(* IEC 61131-3 sources: codesys_asrs/Project_ASRS_CodeSYS, 27 files *)

(* ---- 00_DUT_UDT_MOULE.st ---- *)
// ================================================================
// 00_DUT_UDT_MOULE.st  —  Type utilisateur AS/RS QUADRA 10
// CODESYS V3.5 — DUT (Data Unit Type)
// IMPORTER EN PREMIER dans le projet CODESYS
// ================================================================

TYPE
    UDT_MOULE :
    STRUCT
        ID      : USINT;   // 1=AGADIR 2=IFRANE 3=TANGER 4=RABAT 5=FEZ 0=vide
        OCCUPE  : BOOL;
        RESERVE : BOOL;    // réservé avant prise (évite double allocation)
        RFID_OK : BOOL;    // vérification RFID effectuée sur cet emplacement
    END_STRUCT;
END_TYPE

(* ---- 01_GVL_IO.st ---- *)
// ================================================================
// 01_GVL_IO.st  —  Signaux physiques I/O (GVL nommée "GVL_IO")
// CODESYS V3.5 — Global Variable List
// Sur SoftPLC : pas d'adresse matérielle — simulé via Visualization
//
// Modification v2 — Laser OSSD :
//   ZONE_LIBRE_BTN supprimé → remplacé par OSSD_ZPM + OSSD_PRESSE
//   (Sick S3000 SIL 2 / PLd ISO 13849 — sortie OSSD double canal)
// ================================================================

VAR_GLOBAL
    // ── ENTRÉES CAPTEURS POSITION X ──────────────────────────────
    POS_P0  : BOOL;   // Chariot en P0 (ZPM)
    POS_P1  : BOOL;   // Chariot en P1 (AGADIR)
    POS_P2  : BOOL;   // Chariot en P2 (IFRANE)
    POS_P3  : BOOL;   // Chariot en P3 (TANGER)
    POS_P4  : BOOL;   // Chariot en P4 (RABAT)
    POS_P5  : BOOL;   // Chariot en P5 (FEZ)
    POS_P6  : BOOL;   // Chariot en P6 (Garage)

    // ── ENTRÉES PRÉSENCE CHAMBRES ─────────────────────────────────
    CH1N1   : BOOL;
    CH1N2   : BOOL;
    CH2N1   : BOOL;
    CH2N2   : BOOL;
    CH3N1   : BOOL;
    CH3N2   : BOOL;
    CH4N1   : BOOL;
    CH4N2   : BOOL;
    CH5N1   : BOOL;
    CH5N2   : BOOL;

    // ── ENTRÉES AXE Z ─────────────────────────────────────────────
    CAPTEUR_Z_ZPM       : BOOL;
    CAPTEUR_Z_NIVEAU1   : BOOL;
    CAPTEUR_Z_NIVEAU2   : BOOL;
    CAPTEUR_Z_TRANSPORT : BOOL;

    // ── ENTRÉES SATELLITE ─────────────────────────────────────────
    CAPTEUR_SAT_RETRACTE : BOOL;
    CAPTEUR_SAT_ETENDU   : BOOL;

    // ── ENTRÉES ROTATION ──────────────────────────────────────────
    CAPTEUR_ROT_NORD   : BOOL;
    CAPTEUR_ROT_SUD    : BOOL;
    CAPTEUR_ROT_NEUTRE : BOOL;

    // ── ENTRÉES SÉCURITÉ / ZONE ───────────────────────────────────
    // OSSD : Output Signal Switching Device — Sick S3000 (SIL 2 / PLd)
    // TRUE = zone libre (faisceau non interrompu), FALSE = présence détectée
    OSSD_ZPM              : BOOL;   // Scanner laser zone ZPM P0 (au-dessus de la ZPM)
    OSSD_PRESSE           : BOOL;   // Scanner laser zone presse QUADRA 10
    CAPTEUR_ZONE_OCCUPEE  : BOOL;   // Détecteur de présence (sécurité complémentaire)
    CAPTEUR_CHARGE_CHARIOT: BOOL;

    // ── ENTRÉES RFID ──────────────────────────────────────────────
    RFID_LECTURE_OK : BOOL;
    RFID_ID_LU      : USINT;

    // ── ENTRÉES PRESSE ────────────────────────────────────────────
    PRESSE_ARRETEE      : BOOL;
    PILON_HAUT_OK       : BOOL;
    PILON_BAS_OK        : BOOL;
    MOULE_DEBRIDE       : BOOL;
    MOULE_BRIDE         : BOOL;

    // ── ENTRÉES INTRODUCTEUR ──────────────────────────────────────
    MOULE_SUR_INTRO         : BOOL;
    INTRODUCTEUR_EN_PRESSE  : BOOL;
    INTRODUCTEUR_A_ZPM      : BOOL;
    INTRO_VIDE              : BOOL;

    // ── ENTRÉES COMMANDES OPÉRATEUR (HMI / boutons) ───────────────
    CMD_CM              : BOOL;   // Démarrage changement moule
    CMD_RESET           : BOOL;
    CMD_ACQ_DEF         : BOOL;   // Acquittement défaut
    CMD_HOMING_MANUEL   : BOOL;
    PROLONG_NETTOYAGE_BTN : BOOL; // Demande unique +5 min nettoyage apres alarme T15
    AU_ACTIF            : BOOL;   // Arrêt urgence SW
    MOULE_DEMANDE_HMI   : USINT;  // 1-5
    MODE_AUTO           : BOOL;

    // ── SORTIES AXES ──────────────────────────────────────────────
    CMD_X_AV    : BOOL;
    CMD_X_AR    : BOOL;
    CMD_Z_HAUT  : BOOL;
    CMD_Z_BAS   : BOOL;

    // ── SORTIES SATELLITE ─────────────────────────────────────────
    CMD_SAT_EXT : BOOL;
    CMD_SAT_RET : BOOL;

    // ── SORTIES ROTATION ──────────────────────────────────────────
    CMD_ROT_NORD : BOOL;
    CMD_ROT_SUD  : BOOL;

    // ── SORTIES PRESSE ────────────────────────────────────────────
    CMD_ARRET_PRESSE        : BOOL;
    CMD_DEBRIDAGE           : BOOL;
    CMD_BRIDAGE             : BOOL;
    CMD_AUTORISE_DEMARRAGE  : BOOL;
    CMD_MONTE_PILON         : BOOL;
    CMD_BAISSE_PILON        : BOOL;

    // ── SORTIES INTRODUCTEUR ──────────────────────────────────────
    CMD_INTRO_ENTRE : BOOL;
    CMD_INTRO_SORT  : BOOL;

    // ── SORTIES RFID ──────────────────────────────────────────────
    CMD_RFID_ACTIVER : BOOL;

    // ── SORTIES ENCODEUR / VARIATEUR ──────────────────────────────
    INIT_ENCODEUR_X : BOOL;
    CONSIGNE_POS_X  : WORD;

    // ── SORTIES VOYANTS / BUZZER ──────────────────────────────────
    VOYANT_MACHINE_PRETE    : BOOL;
    VOYANT_CYCLE_EN_COURS   : BOOL;
    VOYANT_DEFAUT           : BOOL;
    VOYANT_INIT_OK          : BOOL;
    VOYANT_NETTOYAGE        : BOOL;
    BUZZER_DEBUT_NETTOYAGE  : BOOL;
    BUZZER_ATTENTE_ZONE_LIBRE : BOOL;
    VOYANT_ATTENTE_ZONE_LIBRE : BOOL;
    VOYANT_NETTOYAGE_TIMEOUT : BOOL;
    VOYANT_NETTOYAGE_MAX     : BOOL;
END_VAR

(* ---- 02_GVL_SIG.st ---- *)
// ================================================================
// 02_GVL_SIG.st  —  Signaux inter-GRAFCETs (GVL nommée "GVL_SIG")
// Équivalent CODESYS de DB_SIG (TIA Portal)
// Point de communication central entre G0-G10
//
// Modification v2 — Laser OSSD + chronos séparés :
//   - Section LASER OSSD ajoutée (Sick S3000)
//   - OSSD_ZONE_LIBRE_AUTO remplace ZONE_LIBRE_BTN comme source de ZONE_CONFIRMEE
//   - Variables chrono chariot / chrono nettoyage séparées
// ================================================================

VAR_GLOBAL
    // ─── SÉCURITÉ (calculé par G1) ───────────────────────────────────
    SECURITES_OK    : BOOL;
    ZONE_CONFIRMEE  : BOOL;   // Géré par FB_LaserSafe — NE PAS écrire depuis HMI directement
    DEFAUT_AXE      : BOOL;
    PERTE_PROFINET  : BOOL;

    // ─── LASER OSSD (Sick S3000 SIL 2 / PLd — géré par FB_LaserSafe) ────
    LASER_ZPM_LIBRE         : BOOL;   // Miroir OSSD_ZPM — zone ZPM libre
    LASER_PRESSE_LIBRE      : BOOL;   // Miroir OSSD_PRESSE — zone presse libre
    OSSD_ZONE_LIBRE_AUTO    : BOOL;   // TRUE après T_ZONE_LIBRE_CONFIRM secondes confirmées
    LASER_MUTING_ACTIF      : BOOL;   // TRUE si CAPTEUR_Z_TRANSPORT — chariot en transit (muting)
    LASER_CONFIRM_EN_COURS  : BOOL;   // Timer de confirmation en cours

    // ─── COMMANDES OPÉRATEUR ─────────────────────────────────────────
    OP_CMD_CM        : BOOL;
    OP_CMD_RESET     : BOOL;
    OP_CMD_ACQ       : BOOL;
    OP_CMD_HOMING    : BOOL;
    OP_MOULE_DEMANDE : USINT;
    OP_MODE_AUTO     : BOOL;
    OP_AU            : BOOL;
    OP_PROLONG_NETTOYAGE : BOOL;

    // ─── G0 ↔ G2 (Homing) ────────────────────────────────────────────
    G2_REQ        : BOOL;
    G2_HOMING_OK  : BOOL;
    G2_DEFAUT     : BOOL;

    // ─── G0 ↔ G3 (Cycle) ─────────────────────────────────────────────
    G3_REQ          : BOOL;
    G3_FIN_CM       : BOOL;
    G3_DEFAUT       : BOOL;
    G3_CODE_DEFAUT  : USINT;

    // ─── G3 ↔ G4 — Axe X ─────────────────────────────────────────────
    G4_REQ   : BOOL;
    G4_CIBLE : USINT;
    G4_DONE  : BOOL;
    G4_ERR   : BOOL;

    // ─── G3 ↔ G5 — Axe Z ─────────────────────────────────────────────
    G5_REQ   : BOOL;
    G5_CIBLE : USINT;
    G5_DONE  : BOOL;
    G5_ERR   : BOOL;

    // ─── G3 ↔ G6 — Rotation ──────────────────────────────────────────
    G6_REQ   : BOOL;
    G6_CIBLE : USINT;
    G6_DONE  : BOOL;
    G6_ERR   : BOOL;

    // ─── G3 ↔ G7 — Satellite ─────────────────────────────────────────
    G7_REQ  : BOOL;
    G7_CMD  : USINT;
    G7_DONE : BOOL;
    G7_ERR  : BOOL;

    // ─── G3 ↔ G8 — RFID ──────────────────────────────────────────────
    G8_REQ        : BOOL;
    G8_ID_ATTENDU : USINT;
    G8_DONE       : BOOL;
    G8_OK         : BOOL;
    G8_ID_LU      : USINT;
    G8_ERR        : BOOL;

    // ─── G3 ↔ G9 — Interface Presse ──────────────────────────────────
    G9_REQ_ARRET      : BOOL;
    G9_REQ_DEBRIDAGE  : BOOL;
    G9_REQ_BRIDAGE    : BOOL;
    G9_REQ_AUTORISER  : BOOL;
    G9_ARRETEE_OK     : BOOL;
    G9_DEBRIDE_OK     : BOOL;
    G9_BRIDE_OK       : BOOL;
    G9_AUTORISE_OK    : BOOL;
    G9_DEFAUT         : BOOL;
    G9_CODE_DEFAUT    : USINT;

    // ─── G3 ↔ G10 — Introducteur ZPM ────────────────────────────────
    G10_REQ_ENTRER : BOOL;
    G10_REQ_SORTIR : BOOL;
    G10_EN_PRESSE  : BOOL;
    G10_A_ZPM      : BOOL;
    G10_DEFAUT     : BOOL;

    // ─── ALARMES ─────────────────────────────────────────────────────
    ALM_STOCK_PLEIN  : BOOL;
    ALM_RFID         : BOOL;
    ALM_DEBRIDAGE    : BOOL;
    ALM_BRIDAGE      : BOOL;
    ALM_PILON        : BOOL;
    ALM_INTRO        : BOOL;
    ALM_AXE_X        : BOOL;
    ALM_AXE_Z        : BOOL;
    ALM_ROTATION     : BOOL;
    ALM_SATELLITE    : BOOL;
    ALM_COMM_PRESSE  : BOOL;
    ALM_ZONE         : BOOL;
    ALM_HOMING       : BOOL;

    // ─── VOYANTS HMI ─────────────────────────────────────────────────
    VYT_MACHINE_PRETE   : BOOL;
    VYT_CYCLE_EN_COURS  : BOOL;
    VYT_DEFAUT          : BOOL;
    VYT_INIT_OK         : BOOL;
    VYT_NETTOYAGE       : BOOL;
    VYT_ATTENTE_ZONE    : BOOL;
    VYT_NETTOYAGE_TIMEOUT : BOOL;

    // ─── NETTOYAGE OPÉRATEUR ─────────────────────────────────────────
    // Surveillance 15 min + prolongation unique 5 min (G3 ET#2 Branche B)
    NETTOYAGE_EN_COURS              : BOOL;
    NETTOYAGE_TIMEOUT               : BOOL;
    NETTOYAGE_PROLONGATION_UTILISEE : BOOL;
    NETTOYAGE_DEPASSEMENT_MAX       : BOOL;

    // ─── ÉTAT SYSTÈME ────────────────────────────────────────────────
    CYCLE_CM_AUTORISE : BOOL;

    // ─── IMAGES I/O (rafraîchies par PLC_PRG avant tout appel FB) ─
    CAPTEUR_POS_X   : ARRAY[0..6] OF BOOL;
    CAPTEUR_PRES_CH : ARRAY[1..5, 1..2] OF BOOL;
END_VAR

(* ---- 03_GVL_MOULES.st ---- *)
// ================================================================
// 03_GVL_MOULES.st  —  Base de données stock moules (GVL "GVL_MOULES")
// Équivalent CODESYS de DB_MOULES (TIA Portal)
// 5 chambres × 2 niveaux = 10 emplacements
// Les valeurs initiales sont chargées par PRG_STARTUP
// ================================================================

VAR_GLOBAL
    // ── Stock physique ────────────────────────────────────────────
    CH : ARRAY[1..5, 1..2] OF UDT_MOULE;   // [chambre 1-5, niveau 1-2]

    // ── État presse et demande ────────────────────────────────────
    MOULE_EN_PRESSE        : USINT;
    MOULE_DEMANDE          : USINT;

    // ── Compteur disponibilité ────────────────────────────────────
    NB_EMPLACEMENTS_LIBRES : USINT;

    // ── Cibles calculées par G3 ───────────────────────────────────
    CIBLE_DEPOT_CH : USINT;
    CIBLE_DEPOT_NV : USINT;
    CIBLE_PRISE_CH : USINT;
    CIBLE_PRISE_NV : USINT;

    // ── Alarme saturation ─────────────────────────────────────────
    ALM_STOCK_PLEIN : BOOL;
END_VAR

(* ---- 04_GVL_SEQ.st ---- *)
// ================================================================
// 04_GVL_SEQ.st  —  État séquence (GVL "GVL_SEQ")
// Équivalent CODESYS de DB_SEQ (TIA Portal)
// Variables RETAIN : survivent au redémarrage (cocher Retain dans CODESYS)
// ================================================================

VAR_GLOBAL
    ETAPE_ACTIVE   : INT;
    CYCLE_EN_COURS : BOOL;
    HOMING_OK      : BOOL;
    DEFAUT_ACTIF   : BOOL;
    CODE_DEFAUT    : USINT;
    // Codes défaut :
    //  1=Timeout arret presse   2=Timeout debridage    3=Timeout bridage
    //  4=Timeout pilon          5=Timeout introducteur 6=Timeout Z
    //  7=Timeout X              8=RFID chambre KO      9=RFID ZPM KO
    // 10=Prise échouée         11=Depot échoue        12=Stock plein
    // 13=Moule introuvable     14=AU pendant cycle    15=Defaut homing
    // 16=Moule presse inconnu  17=Moule demande deja en presse
    // 18=Depassement nettoyage operateur 15+5 min
    // 20=Perte Profinet presse

    // ── Variables RETAIN (cocher "Retain" sur ces variables dans CODESYS)
    CYCLE_INTERROMPU  : BOOL;   // TRUE si coupure pendant cycle
    MOULE_EN_TRANSIT  : BOOL;   // TRUE si moule entre 2 positions
    NB_CYCLES_TOTAL   : DINT;   // compteur cumulé
END_VAR

(* ---- 05_GVL_CFG.st ---- *)
// ================================================================
// 05_GVL_CFG.st  —  Constantes de configuration (GVL "GVL_CFG")
// Équivalent CODESYS de DB_CFG (TIA Portal)
// Positions mécaniques (mm × 10) et timeouts
// ================================================================

VAR_GLOBAL
    // ── Positions Z (unités encoder, 0 = bas) ────────────────────
    Z_ZPM       : INT := 200;
    Z_NIVEAU1   : INT := 450;
    Z_NIVEAU2   : INT := 950;
    Z_TRANSPORT : INT := 1200;

    // ── Positions X (0=P0_ZPM .. 6=P6_Garage) ───────────────────
    X_P0 : INT :=    0;
    X_P1 : INT :=  500;
    X_P2 : INT := 1000;
    X_P3 : INT := 1500;
    X_P4 : INT := 2000;
    X_P5 : INT := 2500;
    X_P6 : INT := 3000;

    // ── Timeouts mouvements et presse ────────────────────────────
    T_ARRET_PRESSE : TIME := T#120S;
    T_DEBRIDAGE    : TIME := T#120S;
    T_BRIDAGE      : TIME := T#120S;
    T_PILON        : TIME := T#120S;
    T_INTRO        : TIME := T#120S;
    T_MVT_Z        : TIME := T#120S;
    T_MVT_X        : TIME := T#120S;
    T_RFID         : TIME := T#120S;
    T_ROTATION     : TIME := T#120S;
    T_SATELLITE    : TIME := T#120S;

    // ── Timeout laser OSSD — confirmation zone libre ──────────────
    // Durée pendant laquelle les deux zones doivent rester libres
    // (OSSD_ZPM=TRUE ET OSSD_PRESSE=TRUE) avant que ZONE_CONFIRMEE soit validée.
    // Norme ISO 13849 / IEC 62061 — délai anti-rebond opérationnel.
    T_ZONE_LIBRE_CONFIRM : TIME := T#10S;
END_VAR

(* ---- 20_GVL_HMI.st ---- *)
// ================================================================
// 20_GVL_HMI.st  —  Variables globales IHM CODESYS Visualization
// GVL nommée "GVL_HMI" dans le projet
// Lier ces variables aux éléments visuels (voir guide 23_CODESYS_HMI_Guide.txt)
// ================================================================

VAR_GLOBAL

    // ── Textes dynamiques (mis à jour par FB_HMI_Controller) ─────
    HMI_MODE_TXT         : STRING(20) := 'HORS SERVICE';
    HMI_ETAPE_G3_TXT     : STRING(40) := '---';
    HMI_MOULE_PRESSE_TXT : STRING(10) := '?';
    HMI_MSG_SYSTEME      : STRING(80) := 'Initialisation...';
    HMI_STOCK_TXT        : ARRAY[1..5, 1..2] OF STRING(10);

    // ── Progression cycle G3 ─────────────────────────────────────
    HMI_G3_ETAPE  : INT   := 0;    // Étape courante 0-15
    HMI_G3_PCT    : REAL  := 0.0;  // Pourcentage 0.0-100.0 (pour BarDisplay)

    // ── Sélecteur moule demandé ───────────────────────────────────
    // Lier à un ComboBox : 0=Choisir 1=MOULE_A 2=MOULE_B 3=MOULE_C 4=MOULE_D 5=MOULE_E
    HMI_SEL_MOULE    : INT  := 0;
    HMI_SEL_MOULE_OK : BOOL := FALSE;

    // ── Chronomètre cycle (format "mm:ss") ───────────────────────
    HMI_TEMPS_CYCLE  : STRING(8) := '00:00';

    // ── Boutons opérateur (lier aux boutons Visualization) ───────
    HMI_BTN_HOMING   : BOOL;   // Démarrer homing
    HMI_BTN_AU       : BOOL;   // Arrêt urgence SW
    HMI_BTN_CMD_CM   : BOOL;   // Démarrer changement moule
    HMI_BTN_ACQ      : BOOL;   // Acquitter défauts
    HMI_BTN_ZONE_OK  : BOOL;   // DIAGNOSTIC ONLY — ne déclenche plus ZONE_CONFIRMEE (laser prime)
    HMI_BTN_PROLONG_NETTOYAGE : BOOL; // Prolongation unique nettoyage +5 min

    // ── Modes dégradés — sélection et injection ───────────────────
    // Combo Box : 0=Aucun 1=D1_StockPlein 2=D2_MouleAbsent
    //             3=D3_TimeoutAxe 4=D4_RFID_KO 5=D5_CycleInterrompu
    //             6=D6_ZoneOccupee 7=D7_PerteProfinet 8=D8_CoupureSecteur
    HMI_FAULT_SEL       : INT := 0;
    HMI_FAULT_DESC      : STRING(100) := 'Sélectionner un scénario...';
    HMI_FAULT_RESULT    : STRING(120) := '';
    HMI_BTN_INJECT      : BOOL;
    HMI_BTN_FAULT_RESET : BOOL;
    HMI_FAULT_ACTIVE    : BOOL;

    // ── Couleurs dynamiques ARGB (mis à jour par FB_HMI_Controller)
    // 16#FF000000 = ARGB (A=opaque toujours à FF)
    // Palette: vert=#FF00C800  rouge=#FFFF3030  orange=#FFFFA500
    //          bleu=#FF1C6EBF  gris=#FF404040   jaune=#FFFFF000
    HMI_COL_MODE      : DWORD := 16#FF404040;
    HMI_COL_FAULT_BTN : DWORD := 16#FF8B0000;   // rouge foncé injecté

    // ── Indicateur alarme globale ─────────────────────────────────
    HMI_ALARME_ACTIVE : BOOL;  // TRUE si au moins 1 alarme

END_VAR

(* ---- 21_FC_MouleIDToStr.st ---- *)
// ================================================================
// 21_FC_MouleIDToStr.st  —  Conversion ID moule (USINT) → nom
// CODESYS V3.5 — FUNCTION
// ================================================================

FUNCTION FC_MouleIDToStr : STRING(10)
VAR_INPUT
    ID : USINT;
END_VAR

CASE ID OF
    0: FC_MouleIDToStr := 'VIDE';
    1: FC_MouleIDToStr := 'MOULE_A';
    2: FC_MouleIDToStr := 'MOULE_B';
    3: FC_MouleIDToStr := 'MOULE_C';
    4: FC_MouleIDToStr := 'MOULE_D';
    5: FC_MouleIDToStr := 'MOULE_E';
ELSE
    FC_MouleIDToStr := '???';
END_CASE;

(* ---- 22_FC_EtapeG3ToStr.st ---- *)
// ================================================================
// 22_FC_EtapeG3ToStr.st  —  Conversion étape G3 (INT) → description
// CODESYS V3.5 — FUNCTION
// ================================================================

FUNCTION FC_EtapeG3ToStr : STRING(35)
VAR_INPUT
    Step : INT;
END_VAR

CASE Step OF
    0 : FC_EtapeG3ToStr := 'REPOS';
    1 : FC_EtapeG3ToStr := 'S01 - Arrêt presse + X→P0';
    2 : FC_EtapeG3ToStr := 'S02 - Rotation NORD';
    3 : FC_EtapeG3ToStr := 'S03 - Satellite étendu ZPM';
    4 : FC_EtapeG3ToStr := 'S04 - Z ZPM - Prise ancien moule';
    5 : FC_EtapeG3ToStr := 'S05 - Satellite rétracté';
    6 : FC_EtapeG3ToStr := 'S06 - Z transport + Rotation 0';
    7 : FC_EtapeG3ToStr := 'S07 - X vers chambre dépôt';
    8 : FC_EtapeG3ToStr := 'S08 - Rotation SUD + Z dépôt';
    9 : FC_EtapeG3ToStr := 'S09 - Satellite - Dépôt moule';
    10: FC_EtapeG3ToStr := 'S10 - X vers chambre prise';
    11: FC_EtapeG3ToStr := 'S11 - Z prise + Vérif. RFID';
    12: FC_EtapeG3ToStr := 'S12 - Satellite - Prise nouveau';
    13: FC_EtapeG3ToStr := 'S13 - Retour P0';
    14: FC_EtapeG3ToStr := 'S14 - RFID ZPM + nettoyage zone';
    15: FC_EtapeG3ToStr := 'S15 - Installation + bridage + P6';
ELSE
    FC_EtapeG3ToStr := 'DEFAUT';
END_CASE;

(* ---- 06_FB_G1_Securite.st ---- *)
// ================================================================
// 06_FB_G1_Securite.st  —  GRAFCET G1 : Sécurité globale
// CODESYS V3.5 — FUNCTION_BLOCK
// Tourne EN PARALLÈLE, permanent, en premier dans PLC_PRG
//
// E1=SECURITES_OK  E2=ARRET_SECURITE  E3=ATTENTE_ACQ
// ================================================================

FUNCTION_BLOCK FB_G1_Securite
VAR
    Step : INT := 1;
END_VAR

VAR_INPUT
END_VAR

VAR_OUTPUT
END_VAR

// ── Corps du FB ──────────────────────────────────────────────────
// ZONE_CONFIRMEE est gérée exclusivement par FB_LaserSafe (OSSD Sick S3000)
// G1 surveille uniquement CAPTEUR_ZONE_OCCUPEE pour alarme immédiate

CASE Step OF

// E1 — SECURITES_OK
1:
    GVL_SIG.SECURITES_OK := TRUE;
    GVL_SIG.ALM_ZONE     := FALSE;

    IF GVL_SIG.OP_AU OR GVL_IO.CAPTEUR_ZONE_OCCUPEE
       OR GVL_SIG.DEFAUT_AXE
       OR GVL_SIG.PERTE_PROFINET THEN
        GVL_IO.CMD_X_AV              := FALSE;
        GVL_IO.CMD_X_AR              := FALSE;
        GVL_IO.CMD_Z_HAUT            := FALSE;
        GVL_IO.CMD_Z_BAS             := FALSE;
        GVL_IO.CMD_SAT_EXT           := FALSE;
        GVL_IO.CMD_SAT_RET           := FALSE;
        GVL_IO.CMD_ROT_NORD          := FALSE;
        GVL_IO.CMD_ROT_SUD           := FALSE;
        GVL_IO.CMD_ARRET_PRESSE      := TRUE;
        GVL_IO.CMD_AUTORISE_DEMARRAGE := FALSE;

        GVL_SIG.SECURITES_OK := FALSE;
        GVL_SIG.ALM_ZONE     := GVL_IO.CAPTEUR_ZONE_OCCUPEE;
        GVL_SIG.VYT_DEFAUT   := TRUE;
        Step := 2;
    END_IF;

// E2 — ARRET_SECURITE
2:
    GVL_IO.CMD_X_AV    := FALSE;
    GVL_IO.CMD_X_AR    := FALSE;
    GVL_IO.CMD_Z_HAUT  := FALSE;
    GVL_IO.CMD_Z_BAS   := FALSE;
    GVL_IO.CMD_SAT_EXT := FALSE;
    GVL_IO.CMD_SAT_RET := FALSE;
    GVL_IO.CMD_ROT_NORD := FALSE;
    GVL_IO.CMD_ROT_SUD  := FALSE;
    Step := 3;

// E3 — ATTENTE_ACQ
3:
    GVL_IO.VOYANT_DEFAUT := TRUE;

    IF NOT GVL_SIG.OP_AU
       AND NOT GVL_IO.CAPTEUR_ZONE_OCCUPEE
       AND NOT GVL_SIG.DEFAUT_AXE
       AND NOT GVL_SIG.PERTE_PROFINET
       AND GVL_SIG.OP_CMD_ACQ THEN
        GVL_SIG.VYT_DEFAUT     := FALSE;
        GVL_IO.VOYANT_DEFAUT   := FALSE;
        GVL_IO.CMD_ARRET_PRESSE := FALSE;
        Step := 1;

    ELSIF GVL_SIG.OP_CMD_ACQ
          AND (GVL_SIG.DEFAUT_AXE OR GVL_SIG.PERTE_PROFINET) THEN
        Step := 2;
    END_IF;

END_CASE;

END_FUNCTION_BLOCK

(* ---- 07_FB_G0_Conduite.st ---- *)
// ================================================================
// 07_FB_G0_Conduite.st  —  GRAFCET G0 : Superviseur modes
// CODESYS V3.5 — FUNCTION_BLOCK
//
// E0=HORS_SERVICE  E1=INIT_SYSTEME  E2=ALARME_REPRISE
// E3=HOMING_EN_COURS  E4=EN_ATTENTE  E5=CYCLE_EN_COURS  E6=DEFAUT_GENERAL
// ================================================================

FUNCTION_BLOCK FB_G0_Conduite
VAR
    Step        : INT := 0;
    StartupDone : BOOL;
END_VAR

CASE Step OF

// E0 — HORS SERVICE
0:
    IF NOT StartupDone THEN
        StartupDone := TRUE;
    END_IF;
    Step := 1;

// E1 — INITIALISATION SYSTÈME
1:
    GVL_SIG.VYT_MACHINE_PRETE := FALSE;
    GVL_SIG.VYT_INIT_OK       := FALSE;
    GVL_SIG.G3_REQ            := FALSE;
    GVL_SIG.G2_REQ            := FALSE;
    GVL_SEQ.HOMING_OK         := FALSE;

    IF GVL_SEQ.CYCLE_INTERROMPU THEN
        GVL_SIG.VYT_DEFAUT := TRUE;
        GVL_SIG.ALM_HOMING := TRUE;
        Step := 2;
    ELSE
        Step := 3;
    END_IF;

// E2 — ALARME REPRISE CYCLE
2:
    GVL_SIG.VYT_DEFAUT := TRUE;
    IF GVL_SIG.OP_CMD_ACQ THEN
        GVL_SIG.VYT_DEFAUT := FALSE;
        GVL_SIG.ALM_HOMING := FALSE;
        Step := 3;
    END_IF;

// E3 — HOMING EN COURS
3:
    GVL_SIG.G2_REQ         := TRUE;
    GVL_SIG.VYT_INIT_OK    := FALSE;
    GVL_SEQ.CYCLE_EN_COURS := FALSE;

    IF GVL_SIG.G2_HOMING_OK THEN
        GVL_SIG.G2_REQ      := FALSE;
        GVL_SEQ.HOMING_OK   := TRUE;
        GVL_SIG.VYT_INIT_OK := TRUE;
        Step := 4;

    ELSIF GVL_SIG.G2_DEFAUT THEN
        GVL_SIG.G2_REQ     := FALSE;
        GVL_SIG.ALM_HOMING := TRUE;
        Step := 6;
    END_IF;

// E4 — EN ATTENTE (machine prête)
4:
    GVL_SIG.VYT_MACHINE_PRETE := TRUE;
    GVL_SIG.CYCLE_CM_AUTORISE :=
        GVL_SIG.OP_CMD_CM
        AND GVL_SEQ.HOMING_OK
        AND GVL_SIG.SECURITES_OK
        AND NOT GVL_SEQ.DEFAUT_ACTIF
        AND NOT GVL_SEQ.CYCLE_EN_COURS
        AND NOT GVL_SIG.OP_AU;

    IF GVL_SIG.OP_CMD_HOMING THEN
        GVL_SIG.VYT_MACHINE_PRETE := FALSE;
        GVL_SEQ.HOMING_OK          := FALSE;
        Step := 3;

    ELSIF GVL_SIG.CYCLE_CM_AUTORISE THEN
        GVL_SIG.VYT_MACHINE_PRETE  := FALSE;
        GVL_SIG.VYT_CYCLE_EN_COURS := TRUE;
        GVL_SEQ.CYCLE_EN_COURS     := TRUE;
        GVL_MOULES.MOULE_DEMANDE   := GVL_SIG.OP_MOULE_DEMANDE;
        GVL_SIG.G3_REQ             := TRUE;
        Step := 5;

    ELSIF GVL_SIG.OP_AU OR GVL_SEQ.DEFAUT_ACTIF THEN
        Step := 6;
    END_IF;

// E5 — CYCLE EN COURS
5:
    IF GVL_SIG.G3_FIN_CM THEN
        GVL_SIG.G3_REQ              := FALSE;
        GVL_SIG.G3_FIN_CM           := FALSE;
        GVL_SEQ.CYCLE_EN_COURS      := FALSE;
        GVL_SIG.VYT_CYCLE_EN_COURS  := FALSE;
        GVL_SEQ.NB_CYCLES_TOTAL     := GVL_SEQ.NB_CYCLES_TOTAL + 1;
        Step := 4;

    ELSIF GVL_SIG.OP_AU OR GVL_SIG.G3_DEFAUT THEN
        GVL_SIG.G3_REQ := FALSE;
        Step := 6;
    END_IF;

// E6 — DEFAUT GENERAL
6:
    GVL_SIG.VYT_DEFAUT         := TRUE;
    GVL_SIG.VYT_MACHINE_PRETE  := FALSE;
    GVL_SIG.VYT_CYCLE_EN_COURS := FALSE;
    GVL_SEQ.CYCLE_EN_COURS     := FALSE;

    IF GVL_SIG.OP_CMD_ACQ
       AND GVL_SIG.OP_CMD_RESET
       AND NOT GVL_SIG.OP_AU
       AND NOT GVL_SEQ.DEFAUT_ACTIF THEN
        GVL_SIG.VYT_DEFAUT  := FALSE;
        GVL_SEQ.HOMING_OK   := FALSE;
        GVL_SIG.ALM_HOMING  := FALSE;
        Step := 3;
    END_IF;

END_CASE;

END_FUNCTION_BLOCK

(* ---- 08_FB_G2_Homing.st ---- *)
// ================================================================
// 08_FB_G2_Homing.st  —  GRAFCET G2 : Référencement axes
// CODESYS V3.5 — FUNCTION_BLOCK
// ORDRE STRICT : Z_TRANSPORT → Sat_Ret → X_P0 → Rot_Neutre → X_P6
//
// E0=ATTENTE  E1=HOMING_Z  E2=HOMING_SAT  E3=HOMING_X
// E4=HOMING_ROT  E5=PARKING  E6=HOMING_OK  E7=DEFAUT
// ================================================================

FUNCTION_BLOCK FB_G2_Homing
VAR
    Step  : INT := 0;
    tmr   : TON;
    tmrIN : BOOL;
END_VAR

tmr(IN := tmrIN, PT := GVL_CFG.T_MVT_X);

CASE Step OF

// E0 — ATTENTE LANCEMENT par G0
0:
    tmrIN := FALSE;
    IF GVL_SIG.G2_REQ THEN
        GVL_SIG.G2_HOMING_OK := FALSE;
        GVL_SIG.G2_DEFAUT    := FALSE;
        Step := 1;
    END_IF;

// E1 — HOMING Z → Z_TRANSPORT
1:
    GVL_IO.CMD_Z_HAUT := TRUE;
    GVL_IO.CMD_Z_BAS  := FALSE;
    tmrIN             := TRUE;
    tmr(IN := tmrIN, PT := GVL_CFG.T_MVT_Z);
    IF GVL_IO.CAPTEUR_Z_TRANSPORT THEN
        GVL_IO.CMD_Z_HAUT := FALSE;
        tmrIN             := FALSE;
        Step              := 2;
    ELSIF tmr.Q THEN
        GVL_IO.CMD_Z_HAUT := FALSE;
        tmrIN             := FALSE;
        Step              := 7;
    END_IF;

// E2 — HOMING SAT → Rétraction satellite
2:
    GVL_IO.CMD_SAT_RET := TRUE;
    GVL_IO.CMD_SAT_EXT := FALSE;
    tmrIN              := TRUE;
    tmr(IN := tmrIN, PT := GVL_CFG.T_SATELLITE);
    IF GVL_IO.CAPTEUR_SAT_RETRACTE THEN
        GVL_IO.CMD_SAT_RET := FALSE;
        tmrIN              := FALSE;
        Step               := 3;
    ELSIF tmr.Q THEN
        GVL_IO.CMD_SAT_RET := FALSE;
        tmrIN              := FALSE;
        Step               := 7;
    END_IF;

// E3 — HOMING X → P0
3:
    GVL_IO.CMD_X_AV := TRUE;
    GVL_IO.CMD_X_AR := FALSE;
    tmrIN           := TRUE;
    tmr(IN := tmrIN, PT := GVL_CFG.T_MVT_X);
    IF GVL_IO.POS_P0 THEN
        GVL_IO.CMD_X_AV         := FALSE;
        GVL_IO.INIT_ENCODEUR_X  := TRUE;
        tmrIN                   := FALSE;
        Step                    := 4;
    ELSIF tmr.Q THEN
        GVL_IO.CMD_X_AV := FALSE;
        tmrIN           := FALSE;
        Step            := 7;
    END_IF;

// E4 — HOMING ROT → Position neutre
4:
    GVL_IO.INIT_ENCODEUR_X := FALSE;
    GVL_IO.CMD_ROT_NORD    := TRUE;
    GVL_IO.CMD_ROT_SUD     := FALSE;
    tmrIN                  := TRUE;
    tmr(IN := tmrIN, PT := GVL_CFG.T_ROTATION);
    IF GVL_IO.CAPTEUR_ROT_NEUTRE THEN
        GVL_IO.CMD_ROT_NORD := FALSE;
        tmrIN               := FALSE;
        Step                := 5;
    ELSIF tmr.Q THEN
        GVL_IO.CMD_ROT_NORD := FALSE;
        tmrIN               := FALSE;
        Step                := 7;
    END_IF;

// E5 — DEPLACEMENT PARKING → P6
5:
    GVL_IO.CMD_X_AR := TRUE;
    GVL_IO.CMD_X_AV := FALSE;
    tmrIN           := TRUE;
    tmr(IN := tmrIN, PT := GVL_CFG.T_MVT_X);
    IF GVL_IO.POS_P6 THEN
        GVL_IO.CMD_X_AR := FALSE;
        tmrIN           := FALSE;
        Step            := 6;
    ELSIF tmr.Q THEN
        GVL_IO.CMD_X_AR := FALSE;
        tmrIN           := FALSE;
        Step            := 7;
    END_IF;

// E6 — HOMING TERMINÉ
6:
    GVL_SIG.G2_HOMING_OK      := TRUE;
    GVL_SEQ.CYCLE_INTERROMPU  := FALSE;
    GVL_SIG.G2_REQ            := FALSE;
    Step := 0;

// E7 — DÉFAUT HOMING
7:
    GVL_SIG.G2_DEFAUT    := TRUE;
    GVL_SEQ.DEFAUT_ACTIF := TRUE;
    GVL_SEQ.CODE_DEFAUT  := 15;
    IF GVL_SIG.OP_CMD_ACQ AND GVL_SIG.OP_CMD_RESET THEN
        GVL_SIG.G2_DEFAUT    := FALSE;
        GVL_SEQ.DEFAUT_ACTIF := FALSE;
        GVL_SEQ.CODE_DEFAUT  := 0;
        Step := 0;
    END_IF;

END_CASE;

END_FUNCTION_BLOCK

(* ---- 09_FB_G4_AxeX.st ---- *)
// ================================================================
// 09_FB_G4_AxeX.st  —  GRAFCET G4 : Axe X (déplacement chariot)
// CODESYS V3.5 — FUNCTION_BLOCK
// RÈGLE ABSOLUE : aucun mouvement X si CAPTEUR_Z_TRANSPORT = FALSE
//
// E0=IMMOBILE  E1=VERIF_Z  E2=ALARME_Z  E3=DEPLACEMENT
// E4=FREINAGE  E5=POSITION_OK  E6=DEFAUT
// ================================================================

FUNCTION_BLOCK FB_G4_AxeX
VAR
    Step  : INT := 0;
    tmr   : TON;
    tmrIN : BOOL;
    Cible : USINT;
END_VAR

tmr(IN := tmrIN, PT := GVL_CFG.T_MVT_X);

CASE Step OF

0: // IMMOBILE — attente requête G3
    GVL_IO.CMD_X_AV   := FALSE;
    GVL_IO.CMD_X_AR   := FALSE;
    GVL_SIG.G4_DONE   := FALSE;
    GVL_SIG.G4_ERR    := FALSE;
    tmrIN             := FALSE;
    IF GVL_SIG.G4_REQ THEN
        Cible := GVL_SIG.G4_CIBLE;
        Step  := 1;
    END_IF;

1: // VÉRIF Z_TRANSPORT — interlock absolu
    IF GVL_IO.CAPTEUR_Z_TRANSPORT THEN
        Step := 3;
    ELSE
        Step := 2;
    END_IF;

2: // ALARME Z NON TRANSPORT
    GVL_SIG.ALM_AXE_X := TRUE;
    IF GVL_IO.CAPTEUR_Z_TRANSPORT THEN
        GVL_SIG.ALM_AXE_X := FALSE;
        Step := 3;
    END_IF;

3: // DÉPLACEMENT X vers cible
    IF GVL_SIG.CAPTEUR_POS_X[Cible] THEN
        Step := 5;
    ELSE
        GVL_IO.CONSIGNE_POS_X := INT_TO_WORD(USINT_TO_INT(Cible));
        GVL_IO.CMD_X_AV       := TRUE;
        GVL_IO.CMD_X_AR       := FALSE;
        tmrIN                 := TRUE;
        Step                  := 4;
    END_IF;

4: // Attente arrivée en position
    IF GVL_SIG.CAPTEUR_POS_X[Cible] THEN
        GVL_IO.CMD_X_AV := FALSE;
        GVL_IO.CMD_X_AR := FALSE;
        tmrIN           := FALSE;
        Step            := 5;
    ELSIF tmr.Q THEN
        GVL_IO.CMD_X_AV       := FALSE;
        GVL_IO.CMD_X_AR       := FALSE;
        tmrIN                 := FALSE;
        GVL_SIG.ALM_AXE_X    := TRUE;
        GVL_SEQ.DEFAUT_ACTIF  := TRUE;
        GVL_SEQ.CODE_DEFAUT   := 7;
        Step := 6;
    END_IF;

5: // POSITION ATTEINTE
    GVL_IO.CMD_X_AV  := FALSE;
    GVL_IO.CMD_X_AR  := FALSE;
    GVL_SIG.G4_DONE  := TRUE;
    GVL_SIG.G4_REQ   := FALSE;
    Step := 0;

6: // DÉFAUT AXE X
    GVL_SIG.G4_ERR    := TRUE;
    GVL_SIG.G4_REQ    := FALSE;
    GVL_SIG.DEFAUT_AXE := TRUE;
    IF GVL_SIG.OP_CMD_ACQ AND GVL_SIG.OP_CMD_RESET THEN
        GVL_SIG.G4_ERR    := FALSE;
        GVL_SIG.ALM_AXE_X := FALSE;
        Step := 0;
    END_IF;

END_CASE;

END_FUNCTION_BLOCK

(* ---- 10_FB_G5_AxeZ.st ---- *)
// ================================================================
// 10_FB_G5_AxeZ.st  —  GRAFCET G5 : Axe Z (hauteur fourches)
// CODESYS V3.5 — FUNCTION_BLOCK
// 4 positions : Z_ZPM(0) Z_NIVEAU1(1) Z_NIVEAU2(2) Z_TRANSPORT(3)
//
// E0=IMMOBILE  E1=MONTEE  E2=DESCENTE  E3=POSITION_OK  E4=DEFAUT
// ================================================================

FUNCTION_BLOCK FB_G5_AxeZ
VAR
    Step  : INT := 0;
    tmr   : TON;
    tmrIN : BOOL;
    Cible : USINT;
END_VAR

tmr(IN := tmrIN, PT := GVL_CFG.T_MVT_Z);

CASE Step OF

0: // IMMOBILE — attente requête G3
    GVL_IO.CMD_Z_HAUT := FALSE;
    GVL_IO.CMD_Z_BAS  := FALSE;
    GVL_SIG.G5_DONE   := FALSE;
    GVL_SIG.G5_ERR    := FALSE;
    tmrIN             := FALSE;
    IF GVL_SIG.G5_REQ THEN
        Cible := GVL_SIG.G5_CIBLE;
        // 0=Z_ZPM  1=Z_NIVEAU1  2=Z_NIVEAU2  3=Z_TRANSPORT
        CASE Cible OF
        0:  // Z_ZPM
            IF GVL_IO.CAPTEUR_Z_ZPM THEN
                Step := 3;
            ELSE
                GVL_IO.CMD_Z_BAS := TRUE;
                tmrIN            := TRUE;
                Step             := 2;
            END_IF;
        1:  // Z_NIVEAU1
            IF GVL_IO.CAPTEUR_Z_NIVEAU1 THEN
                Step := 3;
            ELSIF GVL_IO.CAPTEUR_Z_TRANSPORT OR GVL_IO.CAPTEUR_Z_NIVEAU2 THEN
                GVL_IO.CMD_Z_BAS := TRUE;
                tmrIN            := TRUE;
                Step             := 2;
            ELSE
                GVL_IO.CMD_Z_HAUT := TRUE;
                tmrIN             := TRUE;
                Step              := 1;
            END_IF;
        2:  // Z_NIVEAU2
            IF GVL_IO.CAPTEUR_Z_NIVEAU2 THEN
                Step := 3;
            ELSIF GVL_IO.CAPTEUR_Z_TRANSPORT THEN
                GVL_IO.CMD_Z_BAS := TRUE;
                tmrIN            := TRUE;
                Step             := 2;
            ELSE
                GVL_IO.CMD_Z_HAUT := TRUE;
                tmrIN             := TRUE;
                Step              := 1;
            END_IF;
        3:  // Z_TRANSPORT
            IF GVL_IO.CAPTEUR_Z_TRANSPORT THEN
                Step := 3;
            ELSE
                GVL_IO.CMD_Z_HAUT := TRUE;
                tmrIN             := TRUE;
                Step              := 1;
            END_IF;
        END_CASE;
    END_IF;

1: // MONTÉE en cours
    IF CapteurCibleZ(Cible) THEN
        GVL_IO.CMD_Z_HAUT := FALSE;
        tmrIN             := FALSE;
        Step              := 3;
    ELSIF tmr.Q THEN
        GVL_IO.CMD_Z_HAUT     := FALSE;
        tmrIN                 := FALSE;
        GVL_SIG.ALM_AXE_Z    := TRUE;
        GVL_SEQ.DEFAUT_ACTIF  := TRUE;
        GVL_SEQ.CODE_DEFAUT   := 6;
        Step := 4;
    END_IF;

2: // DESCENTE en cours
    IF CapteurCibleZ(Cible) THEN
        GVL_IO.CMD_Z_BAS := FALSE;
        tmrIN            := FALSE;
        Step             := 3;
    ELSIF tmr.Q THEN
        GVL_IO.CMD_Z_BAS      := FALSE;
        tmrIN                 := FALSE;
        GVL_SIG.ALM_AXE_Z    := TRUE;
        GVL_SEQ.DEFAUT_ACTIF  := TRUE;
        GVL_SEQ.CODE_DEFAUT   := 6;
        Step := 4;
    END_IF;

3: // POSITION ATTEINTE
    GVL_IO.CMD_Z_HAUT := FALSE;
    GVL_IO.CMD_Z_BAS  := FALSE;
    GVL_SIG.G5_DONE   := TRUE;
    GVL_SIG.G5_REQ    := FALSE;
    Step := 0;

4: // DÉFAUT AXE Z
    GVL_SIG.G5_ERR     := TRUE;
    GVL_SIG.G5_REQ     := FALSE;
    GVL_SIG.DEFAUT_AXE := TRUE;
    IF GVL_SIG.OP_CMD_ACQ AND GVL_SIG.OP_CMD_RESET THEN
        GVL_SIG.G5_ERR    := FALSE;
        GVL_SIG.ALM_AXE_Z := FALSE;
        Step := 0;
    END_IF;

END_CASE;

END_FUNCTION_BLOCK

// ── Fonction helper : capteur Z pour la cible demandée ────────────
FUNCTION CapteurCibleZ : BOOL
VAR_INPUT
    Cible : USINT;
END_VAR

CASE Cible OF
0: CapteurCibleZ := GVL_IO.CAPTEUR_Z_ZPM;
1: CapteurCibleZ := GVL_IO.CAPTEUR_Z_NIVEAU1;
2: CapteurCibleZ := GVL_IO.CAPTEUR_Z_NIVEAU2;
3: CapteurCibleZ := GVL_IO.CAPTEUR_Z_TRANSPORT;
ELSE CapteurCibleZ := FALSE;
END_CASE;

END_FUNCTION

(* ---- 11_FB_G6_Rotation.st ---- *)
// ================================================================
// 11_FB_G6_Rotation.st  —  GRAFCET G6 : Rotation plateau
// CODESYS V3.5 — FUNCTION_BLOCK
// 2 positions : NORD=0 (face ZPM/presse)  SUD=1 (face chambres)
//
// E0=REPOS  E1=ROTATION_NORD  E2=ROTATION_SUD
// E3=ORIENTATION_OK  E4=DEFAUT
// ================================================================

FUNCTION_BLOCK FB_G6_Rotation
VAR
    Step  : INT := 0;
    tmr   : TON;
    tmrIN : BOOL;
END_VAR

tmr(IN := tmrIN, PT := GVL_CFG.T_ROTATION);

CASE Step OF

0: // REPOS — attente requête G3
    GVL_IO.CMD_ROT_NORD := FALSE;
    GVL_IO.CMD_ROT_SUD  := FALSE;
    GVL_SIG.G6_DONE     := FALSE;
    GVL_SIG.G6_ERR      := FALSE;
    tmrIN               := FALSE;
    IF GVL_SIG.G6_REQ THEN
        IF GVL_SIG.G6_CIBLE = 0 THEN
            IF GVL_IO.CAPTEUR_ROT_NORD THEN
                Step := 3;
            ELSE
                GVL_IO.CMD_ROT_NORD := TRUE;
                tmrIN               := TRUE;
                Step                := 1;
            END_IF;
        ELSE
            IF GVL_IO.CAPTEUR_ROT_SUD THEN
                Step := 3;
            ELSE
                GVL_IO.CMD_ROT_SUD := TRUE;
                tmrIN              := TRUE;
                Step               := 2;
            END_IF;
        END_IF;
    END_IF;

1: // ROTATION VERS NORD
    IF GVL_IO.CAPTEUR_ROT_NORD THEN
        GVL_IO.CMD_ROT_NORD := FALSE;
        tmrIN               := FALSE;
        Step                := 3;
    ELSIF tmr.Q THEN
        GVL_IO.CMD_ROT_NORD   := FALSE;
        tmrIN                 := FALSE;
        GVL_SIG.ALM_ROTATION  := TRUE;
        GVL_SEQ.DEFAUT_ACTIF  := TRUE;
        GVL_SEQ.CODE_DEFAUT   := 12;
        Step := 4;
    END_IF;

2: // ROTATION VERS SUD
    IF GVL_IO.CAPTEUR_ROT_SUD THEN
        GVL_IO.CMD_ROT_SUD := FALSE;
        tmrIN              := FALSE;
        Step               := 3;
    ELSIF tmr.Q THEN
        GVL_IO.CMD_ROT_SUD    := FALSE;
        tmrIN                 := FALSE;
        GVL_SIG.ALM_ROTATION  := TRUE;
        GVL_SEQ.DEFAUT_ACTIF  := TRUE;
        GVL_SEQ.CODE_DEFAUT   := 12;
        Step := 4;
    END_IF;

3: // ORIENTATION OK
    GVL_IO.CMD_ROT_NORD := FALSE;
    GVL_IO.CMD_ROT_SUD  := FALSE;
    GVL_SIG.G6_DONE     := TRUE;
    GVL_SIG.G6_REQ      := FALSE;
    Step := 0;

4: // DÉFAUT ROTATION
    GVL_SIG.G6_ERR      := TRUE;
    GVL_SIG.G6_REQ      := FALSE;
    GVL_SIG.DEFAUT_AXE  := TRUE;
    IF GVL_SIG.OP_CMD_ACQ AND GVL_SIG.OP_CMD_RESET THEN
        GVL_SIG.G6_ERR       := FALSE;
        GVL_SIG.ALM_ROTATION := FALSE;
        Step := 0;
    END_IF;

END_CASE;

END_FUNCTION_BLOCK

(* ---- 12_FB_G7_Satellite.st ---- *)
// ================================================================
// 12_FB_G7_Satellite.st  —  GRAFCET G7 : Satellite / Fourches
// CODESYS V3.5 — FUNCTION_BLOCK
//
// E0=RETRACTEES  E1=VERIF_AVANT_EXT  E2=EXTENSION
// E3=EXTENSION_OK  E4=RETRACTION  E5=RETRACTEES_OK  E6=DEFAUT
//
// GVL_SIG.G7_CMD : 0=ETENDRE  1=RETRACTER
// ================================================================

FUNCTION_BLOCK FB_G7_Satellite
VAR
    Step  : INT := 0;
    tmr   : TON;
    tmrIN : BOOL;
END_VAR

tmr(IN := tmrIN, PT := GVL_CFG.T_SATELLITE);

CASE Step OF

0: // RETRACTÉES — repos
    GVL_IO.CMD_SAT_EXT := FALSE;
    GVL_IO.CMD_SAT_RET := FALSE;
    GVL_SIG.G7_DONE    := FALSE;
    GVL_SIG.G7_ERR     := FALSE;
    tmrIN              := FALSE;
    IF GVL_SIG.G7_REQ THEN
        IF GVL_SIG.G7_CMD = 0 THEN
            Step := 1;   // Extension demandée
        ELSE
            Step := 4;   // Rétraction demandée
        END_IF;
    END_IF;

1: // VÉRIF AVANT EXTENSION
    IF GVL_IO.CAPTEUR_CHARGE_CHARIOT OR NOT GVL_IO.CAPTEUR_Z_TRANSPORT THEN
        GVL_SIG.G7_ERR := TRUE;
        GVL_SIG.G7_REQ := FALSE;
        Step := 6;
    ELSE
        Step := 2;
    END_IF;

2: // EXTENSION en cours
    GVL_IO.CMD_SAT_EXT := TRUE;
    GVL_IO.CMD_SAT_RET := FALSE;
    tmrIN              := TRUE;
    IF GVL_IO.CAPTEUR_SAT_ETENDU THEN
        GVL_IO.CMD_SAT_EXT := FALSE;
        tmrIN              := FALSE;
        Step               := 3;
    ELSIF tmr.Q THEN
        GVL_IO.CMD_SAT_EXT    := FALSE;
        tmrIN                 := FALSE;
        GVL_SIG.ALM_SATELLITE := TRUE;
        GVL_SEQ.DEFAUT_ACTIF  := TRUE;
        GVL_SEQ.CODE_DEFAUT   := 11;
        Step := 6;
    END_IF;

3: // EXTENSION CONFIRMÉE
    GVL_SIG.G7_DONE := TRUE;
    GVL_SIG.G7_REQ  := FALSE;
    Step := 0;

4: // RÉTRACTION en cours
    GVL_IO.CMD_SAT_RET := TRUE;
    GVL_IO.CMD_SAT_EXT := FALSE;
    tmrIN              := TRUE;
    IF GVL_IO.CAPTEUR_SAT_RETRACTE THEN
        GVL_IO.CMD_SAT_RET := FALSE;
        tmrIN              := FALSE;
        Step               := 5;
    ELSIF tmr.Q THEN
        GVL_IO.CMD_SAT_RET    := FALSE;
        tmrIN                 := FALSE;
        GVL_SIG.ALM_SATELLITE := TRUE;
        GVL_SEQ.DEFAUT_ACTIF  := TRUE;
        GVL_SEQ.CODE_DEFAUT   := 11;
        Step := 6;
    END_IF;

5: // RÉTRACTION CONFIRMÉE
    GVL_SIG.G7_DONE := TRUE;
    GVL_SIG.G7_REQ  := FALSE;
    Step := 0;

6: // DÉFAUT SATELLITE
    GVL_IO.CMD_SAT_EXT    := FALSE;
    GVL_IO.CMD_SAT_RET    := FALSE;
    GVL_SIG.G7_ERR        := TRUE;
    GVL_SIG.G7_REQ        := FALSE;
    GVL_SIG.DEFAUT_AXE    := TRUE;
    IF GVL_SIG.OP_CMD_ACQ AND GVL_SIG.OP_CMD_RESET THEN
        GVL_SIG.G7_ERR        := FALSE;
        GVL_SIG.ALM_SATELLITE := FALSE;
        Step := 0;
    END_IF;

END_CASE;

END_FUNCTION_BLOCK

(* ---- 13_FB_G8_RFID.st ---- *)
// ================================================================
// 13_FB_G8_RFID.st  —  GRAFCET G8 : Lecture RFID
// CODESYS V3.5 — FUNCTION_BLOCK
//
// E0=ATTENTE  E1=LECTURE  E2=COMPARAISON
// E3=RFID_OK  E4=DEFAUT_RFID
// ================================================================

FUNCTION_BLOCK FB_G8_RFID
VAR
    Step  : INT := 0;
    tmr   : TON;
    tmrIN : BOOL;
END_VAR

tmr(IN := tmrIN, PT := GVL_CFG.T_RFID);

CASE Step OF

0: // ATTENTE requête G3
    GVL_IO.CMD_RFID_ACTIVER := FALSE;
    GVL_SIG.G8_DONE         := FALSE;
    GVL_SIG.G8_OK           := FALSE;
    GVL_SIG.G8_ERR          := FALSE;
    GVL_SIG.G8_ID_LU        := 0;
    tmrIN                   := FALSE;
    IF GVL_SIG.G8_REQ THEN
        Step := 1;
    END_IF;

1: // LECTURE RFID
    GVL_IO.CMD_RFID_ACTIVER := TRUE;
    tmrIN                   := TRUE;
    IF GVL_IO.RFID_LECTURE_OK THEN
        GVL_SIG.G8_ID_LU := GVL_IO.RFID_ID_LU;
        tmrIN            := FALSE;
        Step             := 2;
    ELSIF tmr.Q THEN
        GVL_IO.CMD_RFID_ACTIVER := FALSE;
        tmrIN                   := FALSE;
        GVL_SIG.ALM_RFID        := TRUE;
        GVL_SEQ.DEFAUT_ACTIF    := TRUE;
        GVL_SEQ.CODE_DEFAUT     := 8;
        Step := 4;
    END_IF;

2: // COMPARAISON
    GVL_IO.CMD_RFID_ACTIVER := FALSE;
    IF GVL_SIG.G8_ID_LU = GVL_SIG.G8_ID_ATTENDU THEN
        Step := 3;
    ELSE
        GVL_SIG.ALM_RFID      := TRUE;
        GVL_SEQ.DEFAUT_ACTIF  := TRUE;
        GVL_SEQ.CODE_DEFAUT   := 9;
        Step := 4;
    END_IF;

3: // RFID OK
    GVL_SIG.G8_OK   := TRUE;
    GVL_SIG.G8_DONE := TRUE;
    GVL_SIG.G8_REQ  := FALSE;
    Step := 0;

4: // DÉFAUT RFID
    GVL_SIG.G8_OK   := FALSE;
    GVL_SIG.G8_DONE := TRUE;
    GVL_SIG.G8_ERR  := TRUE;
    GVL_SIG.G8_REQ  := FALSE;
    IF NOT GVL_SIG.G8_ERR THEN
        Step := 0;
    END_IF;

END_CASE;

END_FUNCTION_BLOCK

(* ---- 14_FB_G9_Presse.st ---- *)
// ================================================================
// 14_FB_G9_Presse.st  —  GRAFCET G9 : Interface presse QUADRA 10
// CODESYS V3.5 — FUNCTION_BLOCK
//
// Séquence : ARRET → PILON_HAUT → DEBRIDAGE → (cycle chariot)
//            → PILON_BAS → BRIDAGE → AUTORISATION DEMARRAGE
// ================================================================

FUNCTION_BLOCK FB_G9_Presse
VAR
    Step  : INT := 0;
    tmr   : TON;
    tmrIN : BOOL;
END_VAR

tmr(IN := tmrIN, PT := T#1S);

CASE Step OF

// ─── ÉTAT REPOS ──────────────────────────────────────────────
0:
    GVL_IO.CMD_ARRET_PRESSE        := FALSE;
    GVL_IO.CMD_DEBRIDAGE           := FALSE;
    GVL_IO.CMD_BRIDAGE             := FALSE;
    GVL_IO.CMD_AUTORISE_DEMARRAGE  := FALSE;
    GVL_IO.CMD_MONTE_PILON         := FALSE;
    GVL_IO.CMD_BAISSE_PILON        := FALSE;
    GVL_SIG.G9_ARRETEE_OK          := FALSE;
    GVL_SIG.G9_DEBRIDE_OK          := FALSE;
    GVL_SIG.G9_BRIDE_OK            := FALSE;
    GVL_SIG.G9_AUTORISE_OK         := FALSE;
    tmrIN                          := FALSE;
    IF GVL_SIG.G9_REQ_ARRET THEN
        Step := 1;
    END_IF;

// ─── PHASE ARRÊT PRESSE ──────────────────────────────────────
1:
    GVL_IO.CMD_ARRET_PRESSE := TRUE;
    tmrIN                   := TRUE;
    tmr(IN := tmrIN, PT := GVL_CFG.T_ARRET_PRESSE);
    Step := 2;

2:
    IF GVL_IO.PRESSE_ARRETEE THEN
        GVL_IO.CMD_ARRET_PRESSE := FALSE;
        tmrIN                   := FALSE;
        GVL_SIG.G9_ARRETEE_OK  := TRUE;
        Step := 3;
    ELSIF tmr.Q THEN
        GVL_IO.CMD_ARRET_PRESSE  := FALSE;
        tmrIN                    := FALSE;
        GVL_SIG.G9_DEFAUT        := TRUE;
        GVL_SIG.G9_CODE_DEFAUT   := 1;
        GVL_SIG.ALM_COMM_PRESSE  := TRUE;
        Step := 20;
    END_IF;

3: // Monte pilon
    GVL_IO.CMD_MONTE_PILON := TRUE;
    tmrIN                  := TRUE;
    tmr(IN := tmrIN, PT := GVL_CFG.T_PILON);
    Step := 4;

4:
    IF GVL_IO.PILON_HAUT_OK THEN
        GVL_IO.CMD_MONTE_PILON := FALSE;
        tmrIN                  := FALSE;
        IF GVL_SIG.G9_REQ_DEBRIDAGE THEN
            Step := 5;
        END_IF;
    ELSIF tmr.Q THEN
        GVL_IO.CMD_MONTE_PILON   := FALSE;
        tmrIN                    := FALSE;
        GVL_SIG.G9_DEFAUT        := TRUE;
        GVL_SIG.G9_CODE_DEFAUT   := 4;
        GVL_SIG.ALM_PILON        := TRUE;
        Step := 20;
    END_IF;

5: // Débridage
    GVL_IO.CMD_DEBRIDAGE := TRUE;
    tmrIN                := TRUE;
    tmr(IN := tmrIN, PT := GVL_CFG.T_DEBRIDAGE);
    Step := 6;

6:
    IF GVL_IO.MOULE_DEBRIDE THEN
        GVL_IO.CMD_DEBRIDAGE     := FALSE;
        tmrIN                    := FALSE;
        GVL_SIG.G9_DEBRIDE_OK    := TRUE;
        Step := 7;
    ELSIF tmr.Q THEN
        GVL_IO.CMD_DEBRIDAGE     := FALSE;
        tmrIN                    := FALSE;
        GVL_SIG.ALM_DEBRIDAGE    := TRUE;
        Step := 15;   // ROLLBACK
    END_IF;

7: // ATTENTE commande bridage
    IF GVL_SIG.G9_REQ_BRIDAGE THEN
        Step := 8;
    END_IF;

// ─── PHASE BRIDAGE ───────────────────────────────────────────
8: // Baisse pilon
    GVL_IO.CMD_BAISSE_PILON := TRUE;
    tmrIN                   := TRUE;
    tmr(IN := tmrIN, PT := GVL_CFG.T_PILON);
    Step := 9;

9:
    IF GVL_IO.PILON_BAS_OK AND GVL_IO.MOULE_SUR_INTRO AND GVL_IO.INTRODUCTEUR_A_ZPM THEN
        GVL_IO.CMD_BAISSE_PILON := FALSE;
        tmrIN                   := FALSE;
        Step := 10;
    ELSIF tmr.Q THEN
        GVL_IO.CMD_BAISSE_PILON  := FALSE;
        tmrIN                    := FALSE;
        GVL_SIG.G9_DEFAUT        := TRUE;
        GVL_SIG.G9_CODE_DEFAUT   := 4;
        GVL_SIG.ALM_PILON        := TRUE;
        Step := 20;
    END_IF;

10: // Bridage
    GVL_IO.CMD_BRIDAGE := TRUE;
    tmrIN              := TRUE;
    tmr(IN := tmrIN, PT := GVL_CFG.T_BRIDAGE);
    Step := 11;

11:
    IF GVL_IO.MOULE_BRIDE THEN
        GVL_IO.CMD_BRIDAGE     := FALSE;
        tmrIN                  := FALSE;
        GVL_SIG.G9_BRIDE_OK    := TRUE;
        Step := 12;
    ELSIF tmr.Q THEN
        GVL_IO.CMD_BRIDAGE       := FALSE;
        tmrIN                    := FALSE;
        GVL_SIG.G9_DEFAUT        := TRUE;
        GVL_SIG.G9_CODE_DEFAUT   := 3;
        GVL_SIG.ALM_BRIDAGE      := TRUE;
        Step := 20;
    END_IF;

12: // ATTENTE autorisation
    IF GVL_SIG.G9_REQ_AUTORISER THEN
        Step := 13;
    END_IF;

13:
    IF GVL_IO.INTRO_VIDE AND GVL_IO.INTRODUCTEUR_A_ZPM THEN
        GVL_IO.CMD_AUTORISE_DEMARRAGE := TRUE;
        Step := 14;
    ELSE
        GVL_SIG.G9_DEFAUT      := TRUE;
        GVL_SIG.G9_CODE_DEFAUT := 5;
        Step := 20;
    END_IF;

14: // AUTORISATION ENVOYÉE
    GVL_SIG.G9_AUTORISE_OK     := TRUE;
    GVL_SIG.G9_REQ_ARRET       := FALSE;
    GVL_SIG.G9_REQ_DEBRIDAGE   := FALSE;
    GVL_SIG.G9_REQ_BRIDAGE     := FALSE;
    GVL_SIG.G9_REQ_AUTORISER   := FALSE;
    Step := 0;

// ─── ROLLBACK DÉBRIDAGE ÉCHOUÉ ───────────────────────────────
15:
    GVL_IO.CMD_BAISSE_PILON := TRUE;
    tmrIN                   := TRUE;
    tmr(IN := tmrIN, PT := GVL_CFG.T_PILON);
    Step := 16;

16:
    IF GVL_IO.PILON_BAS_OK OR tmr.Q THEN
        GVL_IO.CMD_BAISSE_PILON        := FALSE;
        tmrIN                          := FALSE;
        GVL_IO.CMD_AUTORISE_DEMARRAGE  := TRUE;
        GVL_SIG.G9_DEFAUT              := TRUE;
        GVL_SIG.G9_CODE_DEFAUT         := 2;
        Step := 17;
    END_IF;

17:
    IF NOT GVL_IO.PRESSE_ARRETEE THEN
        GVL_IO.CMD_AUTORISE_DEMARRAGE := FALSE;
        Step := 0;
    END_IF;

// ─── DÉFAUT GÉNÉRAL G9 ───────────────────────────────────────
20:
    GVL_IO.CMD_ARRET_PRESSE        := FALSE;
    GVL_IO.CMD_DEBRIDAGE           := FALSE;
    GVL_IO.CMD_BRIDAGE             := FALSE;
    GVL_IO.CMD_MONTE_PILON         := FALSE;
    GVL_IO.CMD_BAISSE_PILON        := FALSE;
    GVL_IO.CMD_AUTORISE_DEMARRAGE  := FALSE;
    IF GVL_SIG.OP_CMD_ACQ AND GVL_SIG.OP_CMD_RESET THEN
        GVL_SIG.G9_DEFAUT        := FALSE;
        GVL_SIG.G9_CODE_DEFAUT   := 0;
        GVL_SIG.ALM_COMM_PRESSE  := FALSE;
        GVL_SIG.ALM_PILON        := FALSE;
        GVL_SIG.ALM_DEBRIDAGE    := FALSE;
        GVL_SIG.ALM_BRIDAGE      := FALSE;
        Step := 0;
    END_IF;

END_CASE;

END_FUNCTION_BLOCK

(* ---- 15_FB_G10_Intro.st ---- *)
// ================================================================
// 15_FB_G10_Intro.st  —  GRAFCET G10 : Introducteur ZPM
// CODESYS V3.5 — FUNCTION_BLOCK
//
// SÉCURITÉ : Entrée en presse UNIQUEMENT si PILON_HAUT_OK = TRUE
//
// E0=A_ZPM  E1=VERIF_ENTREE  E2=INTRO_EN_COURS
// E3=EN_PRESSE  E4=RETRAIT_EN_COURS  E5=REVENU_ZPM  E6=DEFAUT
// ================================================================

FUNCTION_BLOCK FB_G10_Intro
VAR
    Step  : INT := 0;
    tmr   : TON;
    tmrIN : BOOL;
END_VAR

tmr(IN := tmrIN, PT := GVL_CFG.T_INTRO);

CASE Step OF

0: // À ZPM — état initial
    GVL_IO.CMD_INTRO_ENTRE  := FALSE;
    GVL_IO.CMD_INTRO_SORT   := FALSE;
    GVL_SIG.G10_DEFAUT      := FALSE;
    GVL_SIG.G10_EN_PRESSE   := FALSE;
    GVL_SIG.G10_A_ZPM       := TRUE;
    tmrIN                   := FALSE;
    IF GVL_SIG.G10_REQ_ENTRER THEN
        GVL_SIG.G10_A_ZPM := FALSE;
        Step := 1;
    END_IF;

1: // VÉRIFICATION SÉCURITÉ
    IF NOT GVL_IO.PILON_HAUT_OK THEN
        GVL_SIG.G10_DEFAUT    := TRUE;
        GVL_SEQ.DEFAUT_ACTIF  := TRUE;
        GVL_SEQ.CODE_DEFAUT   := 5;
        GVL_SIG.ALM_INTRO     := TRUE;
        Step := 6;
    ELSE
        GVL_IO.CMD_INTRO_ENTRE := TRUE;
        tmrIN                  := TRUE;
        Step                   := 2;
    END_IF;

2: // INTRODUCTION EN COURS
    IF GVL_IO.INTRODUCTEUR_EN_PRESSE THEN
        GVL_IO.CMD_INTRO_ENTRE  := FALSE;
        tmrIN                   := FALSE;
        GVL_SIG.G10_EN_PRESSE   := TRUE;
        Step := 3;
    ELSIF tmr.Q THEN
        GVL_IO.CMD_INTRO_ENTRE := FALSE;
        tmrIN                  := FALSE;
        GVL_SIG.ALM_INTRO      := TRUE;
        GVL_SEQ.DEFAUT_ACTIF   := TRUE;
        GVL_SEQ.CODE_DEFAUT    := 5;
        Step := 6;
    END_IF;

3: // EN PRESSE — attente commande retrait
    IF GVL_SIG.G10_REQ_SORTIR THEN
        GVL_SIG.G10_EN_PRESSE := FALSE;
        GVL_IO.CMD_INTRO_SORT  := TRUE;
        tmrIN                  := TRUE;
        Step                   := 4;
    END_IF;

4: // RETRAIT EN COURS
    IF GVL_IO.INTRODUCTEUR_A_ZPM THEN
        GVL_IO.CMD_INTRO_SORT := FALSE;
        tmrIN                 := FALSE;
        GVL_SIG.G10_A_ZPM    := TRUE;
        Step                  := 5;
    ELSIF tmr.Q THEN
        GVL_IO.CMD_INTRO_SORT  := FALSE;
        tmrIN                  := FALSE;
        GVL_SIG.ALM_INTRO      := TRUE;
        GVL_SEQ.DEFAUT_ACTIF   := TRUE;
        GVL_SEQ.CODE_DEFAUT    := 5;
        Step := 6;
    END_IF;

5: // REVENU À ZPM
    GVL_SIG.G10_REQ_ENTRER := FALSE;
    GVL_SIG.G10_REQ_SORTIR := FALSE;
    Step := 0;

6: // DÉFAUT INTRODUCTEUR
    GVL_IO.CMD_INTRO_ENTRE  := FALSE;
    GVL_IO.CMD_INTRO_SORT   := FALSE;
    GVL_SIG.G10_DEFAUT      := TRUE;
    IF GVL_SIG.OP_CMD_ACQ AND GVL_SIG.OP_CMD_RESET THEN
        GVL_SIG.G10_DEFAUT      := FALSE;
        GVL_SIG.G10_REQ_ENTRER  := FALSE;
        GVL_SIG.G10_REQ_SORTIR  := FALSE;
        GVL_SIG.ALM_INTRO       := FALSE;
        Step := 0;
    END_IF;

END_CASE;

END_FUNCTION_BLOCK

(* ---- 16_FB_G3_Cycle.st ---- *)
// ================================================================
// 16_FB_G3_Cycle.st  —  GRAFCET G3 : Coordinateur cycle AS/RS
// CODESYS V3.5 — FUNCTION_BLOCK
// Chef d'orchestre — active G4..G10 via GVL_SIG
//
// 3 DIVERGENCES ET :
//   ET#1 : retrait introducteur ‖ chariot → P0
//   ET#2 : stockage+RFID+prise ‖ nettoyage opérateurs
//   ET#3 : autorisation presse ‖ retour garage
// ================================================================

FUNCTION_BLOCK FB_G3_Cycle
VAR
    Step       : INT := 0;
    SubA       : INT;
    SubB       : INT;
    BrA_Done   : BOOL;
    BrB_Done   : BOOL;
    i          : INT;
    j          : INT;
    DepotFound : BOOL;
    PriseFound : BOOL;
    NvZ        : USINT;
    T_Nettoyage15 : TON;
    T_Prolong5   : TON;
    NettoyageTimerEnable : BOOL;
    ProlongTimerEnable   : BOOL;
END_VAR

T_Nettoyage15(IN := NettoyageTimerEnable AND NOT GVL_SIG.ZONE_CONFIRMEE, PT := T#15m);
T_Prolong5(IN := ProlongTimerEnable AND NOT GVL_SIG.ZONE_CONFIRMEE, PT := T#5m);

// ── Surveillance AU pendant cycle (priorité absolue) ──────────
IF GVL_SIG.OP_AU AND Step > 0 AND Step < 200 THEN
    GVL_SIG.G3_DEFAUT      := TRUE;
    GVL_SIG.G3_CODE_DEFAUT := 14;
    GVL_SEQ.DEFAUT_ACTIF   := TRUE;
    GVL_SEQ.CODE_DEFAUT    := 14;
    GVL_SIG.G4_REQ         := FALSE;
    GVL_SIG.G5_REQ         := FALSE;
    GVL_SIG.G6_REQ         := FALSE;
    GVL_SIG.G7_REQ         := FALSE;
    GVL_SIG.G8_REQ         := FALSE;
    GVL_SIG.G9_REQ_ARRET     := FALSE;
    GVL_SIG.G10_REQ_ENTRER   := FALSE;
    GVL_SIG.G10_REQ_SORTIR   := FALSE;
    GVL_SIG.VYT_CYCLE_EN_COURS := FALSE;
    Step := 0;
    RETURN;
END_IF;

CASE Step OF

// ════════════════════════════════════════════════════════════
// PHASE 0 — IDLE
// ════════════════════════════════════════════════════════════
0:
    GVL_SIG.G3_FIN_CM          := FALSE;
    GVL_SIG.G3_DEFAUT          := FALSE;
    GVL_SIG.G3_CODE_DEFAUT     := 0;
    GVL_SIG.VYT_CYCLE_EN_COURS := FALSE;
    GVL_SIG.G9_ARRETEE_OK      := FALSE;
    GVL_SIG.G9_DEBRIDE_OK      := FALSE;
    GVL_SIG.G9_BRIDE_OK        := FALSE;
    GVL_SIG.G9_AUTORISE_OK     := FALSE;
    GVL_SIG.G10_EN_PRESSE      := FALSE;
    GVL_SIG.G10_A_ZPM          := FALSE;
    NettoyageTimerEnable       := FALSE;
    ProlongTimerEnable         := FALSE;
    GVL_SIG.NETTOYAGE_EN_COURS := FALSE;
    GVL_SIG.NETTOYAGE_TIMEOUT  := FALSE;
    GVL_SIG.NETTOYAGE_PROLONGATION_UTILISEE := FALSE;
    GVL_SIG.NETTOYAGE_DEPASSEMENT_MAX := FALSE;
    GVL_SIG.VYT_NETTOYAGE_TIMEOUT := FALSE;
    GVL_IO.VOYANT_NETTOYAGE_TIMEOUT := FALSE;
    GVL_IO.VOYANT_NETTOYAGE_MAX := FALSE;
    GVL_IO.BUZZER_ATTENTE_ZONE_LIBRE := FALSE;
    IF GVL_SIG.G3_REQ THEN
        DepotFound := FALSE;
        PriseFound := FALSE;
        IF GVL_MOULES.MOULE_EN_PRESSE = 0 THEN
            GVL_SIG.G3_CODE_DEFAUT := 16;
            Step := 200;
        ELSIF GVL_MOULES.MOULE_DEMANDE = 0 THEN
            GVL_SIG.G3_CODE_DEFAUT := 13;
            Step := 200;
        ELSIF GVL_MOULES.MOULE_DEMANDE = GVL_MOULES.MOULE_EN_PRESSE THEN
            GVL_SIG.G3_CODE_DEFAUT := 17;
            Step := 200;
        ELSE
            Step := 1;
        END_IF;
    END_IF;

1: // Recherche slot dépôt
    DepotFound := FALSE;
    FOR i := 1 TO 5 BY 1 DO
        IF NOT DepotFound THEN
            FOR j := 1 TO 2 BY 1 DO
                IF NOT DepotFound
                   AND NOT GVL_MOULES.CH[i, j].OCCUPE
                   AND NOT GVL_MOULES.CH[i, j].RESERVE THEN
                    GVL_MOULES.CIBLE_DEPOT_CH := INT_TO_USINT(i);
                    GVL_MOULES.CIBLE_DEPOT_NV := INT_TO_USINT(j);
                    GVL_MOULES.CH[i, j].RESERVE := TRUE;
                    DepotFound := TRUE;
                END_IF;
            END_FOR;
        END_IF;
    END_FOR;
    IF DepotFound THEN
        Step := 2;
    ELSE
        GVL_MOULES.ALM_STOCK_PLEIN := TRUE;
        GVL_SIG.ALM_STOCK_PLEIN   := TRUE;
        GVL_SIG.G3_CODE_DEFAUT    := 12;
        Step := 200;
    END_IF;

2: // Recherche slot prise
    PriseFound := FALSE;
    FOR i := 1 TO 5 BY 1 DO
        IF NOT PriseFound THEN
            FOR j := 1 TO 2 BY 1 DO
                IF NOT PriseFound
                   AND GVL_MOULES.CH[i, j].OCCUPE
                   AND GVL_MOULES.CH[i, j].ID = GVL_MOULES.MOULE_DEMANDE THEN
                    GVL_MOULES.CIBLE_PRISE_CH := INT_TO_USINT(i);
                    GVL_MOULES.CIBLE_PRISE_NV := INT_TO_USINT(j);
                    PriseFound := TRUE;
                END_IF;
            END_FOR;
        END_IF;
    END_FOR;
    IF PriseFound THEN
        GVL_SIG.VYT_CYCLE_EN_COURS := TRUE;
        Step := 3;
    ELSE
        GVL_MOULES.CH[GVL_MOULES.CIBLE_DEPOT_CH, GVL_MOULES.CIBLE_DEPOT_NV].RESERVE := FALSE;
        GVL_SIG.G3_CODE_DEFAUT := 13;
        Step := 200;
    END_IF;

3:
    GVL_SEQ.CYCLE_INTERROMPU := TRUE;
    GVL_SEQ.CYCLE_EN_COURS   := TRUE;

// ════════════════════════════════════════════════════════════
// PHASE 1 — Arrêt presse + débridage
// ════════════════════════════════════════════════════════════
10:
    GVL_SIG.G9_REQ_ARRET   := TRUE;
    GVL_SIG.G10_REQ_ENTRER := TRUE;
    Step := 11;

11:
    IF GVL_SIG.G9_ARRETEE_OK THEN
        GVL_SIG.G9_REQ_DEBRIDAGE := TRUE;
        Step := 12;
    ELSIF GVL_SIG.G9_DEFAUT THEN
        Step := 200;
    END_IF;

12:
    IF GVL_SIG.G9_DEBRIDE_OK THEN
        Step := 13;
    ELSIF GVL_SIG.G9_DEFAUT THEN
        Step := 200;
    END_IF;

// ════════════════════════════════════════════════════════════
// DIVERGENCE ET#1 — Retrait introducteur ‖ Chariot → P0
// ════════════════════════════════════════════════════════════
13:
    BrA_Done := FALSE;
    BrB_Done := FALSE;
    SubA     := 0;
    SubB     := 0;
    Step     := 14;

14:
    IF NOT BrA_Done THEN
        CASE SubA OF
        0:  GVL_SIG.G10_REQ_SORTIR := TRUE;
            SubA := 1;
        1:  IF GVL_SIG.G10_A_ZPM THEN
                BrA_Done := TRUE;
            ELSIF GVL_SIG.G10_DEFAUT THEN
                GVL_SIG.G3_CODE_DEFAUT := 5;
                Step := 200;
            END_IF;
        END_CASE;
    END_IF;

    IF NOT BrB_Done THEN
        CASE SubB OF
        0:  GVL_SIG.G4_REQ   := TRUE;
            GVL_SIG.G4_CIBLE := 0;
            SubB := 1;
        1:  IF GVL_SIG.G4_DONE THEN
                GVL_SIG.G4_DONE := FALSE;
                BrB_Done := TRUE;
            ELSIF GVL_SIG.G4_ERR THEN
                GVL_SIG.G4_ERR := FALSE;
                GVL_SIG.G3_CODE_DEFAUT := 7;
                Step := 200;
            END_IF;
        END_CASE;
    END_IF;

    IF BrA_Done AND BrB_Done THEN
        GVL_SIG.G10_REQ_ENTRER := FALSE;
        GVL_SIG.G10_REQ_SORTIR := FALSE;
        Step := 15;
    END_IF;

// ════════════════════════════════════════════════════════════
// PHASE 2 — Transfert moule : introducteur → chariot
// ════════════════════════════════════════════════════════════
15:
    IF NOT GVL_IO.MOULE_SUR_INTRO THEN
        GVL_SIG.G3_CODE_DEFAUT := 13;
        Step := 200;
    ELSE
        Step := 16;
    END_IF;

16:
    GVL_SIG.G6_REQ   := TRUE;
    GVL_SIG.G6_CIBLE := 0;  // NORD
    Step := 17;

17:
    IF GVL_SIG.G6_DONE THEN
        GVL_SIG.G6_DONE := FALSE;
        Step := 18;
    ELSIF GVL_SIG.G6_ERR THEN
        GVL_SIG.G6_ERR         := FALSE;
        GVL_SIG.G3_CODE_DEFAUT := 11;
        Step := 200;
    END_IF;

18:
    GVL_SIG.G5_REQ   := TRUE;
    GVL_SIG.G5_CIBLE := 0;  // Z_ZPM
    Step := 19;

19:
    IF GVL_SIG.G5_DONE THEN
        GVL_SIG.G5_DONE := FALSE;
        Step := 20;
    ELSIF GVL_SIG.G5_ERR THEN
        GVL_SIG.G5_ERR         := FALSE;
        GVL_SIG.G3_CODE_DEFAUT := 6;
        Step := 200;
    END_IF;

20:
    GVL_SIG.G7_REQ := TRUE;
    GVL_SIG.G7_CMD := 0;  // ETENDRE
    Step := 21;

21:
    IF GVL_SIG.G7_DONE THEN
        GVL_SIG.G7_DONE := FALSE;
        Step := 22;
    ELSIF GVL_SIG.G7_ERR THEN
        GVL_SIG.G7_ERR         := FALSE;
        GVL_SIG.G3_CODE_DEFAUT := 11;
        Step := 200;
    END_IF;

22:
    GVL_SIG.G5_REQ   := TRUE;
    GVL_SIG.G5_CIBLE := 3;  // Z_TRANSPORT
    Step := 23;

23:
    IF GVL_SIG.G5_DONE THEN
        GVL_SIG.G5_DONE := FALSE;
        IF NOT GVL_IO.CAPTEUR_CHARGE_CHARIOT THEN
            GVL_SIG.G3_CODE_DEFAUT := 10;
            Step := 200;
        ELSE
            Step := 24;
        END_IF;
    ELSIF GVL_SIG.G5_ERR THEN
        GVL_SIG.G5_ERR         := FALSE;
        GVL_SIG.G3_CODE_DEFAUT := 6;
        Step := 200;
    END_IF;

24:
    GVL_SIG.G7_REQ := TRUE;
    GVL_SIG.G7_CMD := 1;  // RETRACTER
    Step := 25;

25:
    IF GVL_SIG.G7_DONE THEN
        GVL_SIG.G7_DONE := FALSE;
        Step := 26;
    ELSIF GVL_SIG.G7_ERR THEN
        GVL_SIG.G7_ERR         := FALSE;
        GVL_SIG.G3_CODE_DEFAUT := 11;
        Step := 201;
    END_IF;

// ════════════════════════════════════════════════════════════
// DIVERGENCE ET#2 — Stockage+RFID+Prise ‖ Nettoyage
// ════════════════════════════════════════════════════════════
26:
    BrA_Done := FALSE;
    BrB_Done := FALSE;
    SubA     := 0;
    SubB     := 0;
    NettoyageTimerEnable := FALSE;
    ProlongTimerEnable := FALSE;
    GVL_SIG.NETTOYAGE_EN_COURS := FALSE;
    GVL_SIG.NETTOYAGE_TIMEOUT := FALSE;
    GVL_SIG.NETTOYAGE_PROLONGATION_UTILISEE := FALSE;
    GVL_SIG.NETTOYAGE_DEPASSEMENT_MAX := FALSE;
    GVL_SIG.VYT_NETTOYAGE_TIMEOUT := FALSE;
    GVL_IO.VOYANT_NETTOYAGE_TIMEOUT := FALSE;
    GVL_IO.VOYANT_NETTOYAGE_MAX := FALSE;
    GVL_IO.BUZZER_ATTENTE_ZONE_LIBRE := FALSE;
    // Réinitialise la validation laser pour forcer une nouvelle confirmation 10s
    // sans ce reset, le 2ème cycle validerait immédiatement si ZONE_CONFIRMEE
    // était encore TRUE depuis le cycle précédent
    GVL_SIG.ZONE_CONFIRMEE    := FALSE;
    GVL_SIG.OSSD_ZONE_LIBRE_AUTO := FALSE;
    Step     := 27;

27: // ET#2
    IF NOT BrA_Done THEN
        CASE SubA OF
        0:  GVL_SIG.G4_REQ   := TRUE;
            GVL_SIG.G4_CIBLE := GVL_MOULES.CIBLE_DEPOT_CH;
            SubA := 1;
        1:  IF GVL_SIG.G4_DONE THEN
                GVL_SIG.G4_DONE := FALSE; SubA := 2;
            ELSIF GVL_SIG.G4_ERR THEN
                GVL_SIG.G4_ERR := FALSE;
                GVL_SIG.G3_CODE_DEFAUT := 7; Step := 201; END_IF;
        2:  GVL_SIG.G6_REQ   := TRUE;
            GVL_SIG.G6_CIBLE := 1; // SUD
            SubA := 3;
        3:  IF GVL_SIG.G6_DONE THEN
                GVL_SIG.G6_DONE := FALSE; SubA := 4;
            ELSIF GVL_SIG.G6_ERR THEN
                GVL_SIG.G6_ERR := FALSE;
                GVL_SIG.G3_CODE_DEFAUT := 11; Step := 201; END_IF;
        4:  GVL_SIG.G7_REQ := TRUE;
            GVL_SIG.G7_CMD := 0; // EXT
            SubA := 5;
        5:  IF GVL_SIG.G7_DONE THEN
                GVL_SIG.G7_DONE := FALSE; SubA := 6;
            ELSIF GVL_SIG.G7_ERR THEN
                GVL_SIG.G7_ERR := FALSE;
                GVL_SIG.G3_CODE_DEFAUT := 11; Step := 201; END_IF;
        6:  GVL_SIG.G5_REQ   := TRUE;
            GVL_SIG.G5_CIBLE := GVL_MOULES.CIBLE_DEPOT_NV;
            SubA := 7;
        7:  IF GVL_SIG.G5_DONE THEN
                GVL_SIG.G5_DONE := FALSE; SubA := 8;
            ELSIF GVL_SIG.G5_ERR THEN
                GVL_SIG.G5_ERR := FALSE;
                GVL_SIG.G3_CODE_DEFAUT := 6; Step := 201; END_IF;
        8:  GVL_SIG.G7_REQ := TRUE;
            GVL_SIG.G7_CMD := 1; // RET
            SubA := 9;
        9:  IF GVL_SIG.G7_DONE THEN
                GVL_SIG.G7_DONE := FALSE;
                IF NOT GVL_SIG.CAPTEUR_PRES_CH[GVL_MOULES.CIBLE_DEPOT_CH,
                                               GVL_MOULES.CIBLE_DEPOT_NV] THEN
                    GVL_SIG.G3_CODE_DEFAUT := 11; Step := 202;
                ELSE
                    GVL_MOULES.CH[GVL_MOULES.CIBLE_DEPOT_CH,
                                  GVL_MOULES.CIBLE_DEPOT_NV].OCCUPE  := TRUE;
                    GVL_MOULES.CH[GVL_MOULES.CIBLE_DEPOT_CH,
                                  GVL_MOULES.CIBLE_DEPOT_NV].ID      := GVL_MOULES.MOULE_EN_PRESSE;
                    GVL_MOULES.CH[GVL_MOULES.CIBLE_DEPOT_CH,
                                  GVL_MOULES.CIBLE_DEPOT_NV].RESERVE := FALSE;
                    IF GVL_MOULES.NB_EMPLACEMENTS_LIBRES > 0 THEN
                        GVL_MOULES.NB_EMPLACEMENTS_LIBRES :=
                            GVL_MOULES.NB_EMPLACEMENTS_LIBRES - 1;
                    END_IF;
                    SubA := 10;
                END_IF;
            ELSIF GVL_SIG.G7_ERR THEN
                GVL_SIG.G7_ERR := FALSE;
                GVL_SIG.G3_CODE_DEFAUT := 11; Step := 202; END_IF;
        10: GVL_SIG.G5_REQ   := TRUE;
            GVL_SIG.G5_CIBLE := 3; // Z_TRANSPORT
            SubA := 11;
        11: IF GVL_SIG.G5_DONE THEN
                GVL_SIG.G5_DONE := FALSE; SubA := 12;
            ELSIF GVL_SIG.G5_ERR THEN
                GVL_SIG.G5_ERR := FALSE;
                GVL_SIG.G3_CODE_DEFAUT := 6; Step := 202; END_IF;
        12: GVL_SIG.G4_REQ   := TRUE;
            GVL_SIG.G4_CIBLE := GVL_MOULES.CIBLE_PRISE_CH;
            SubA := 13;
        13: IF GVL_SIG.G4_DONE THEN
                GVL_SIG.G4_DONE := FALSE; SubA := 14;
            ELSIF GVL_SIG.G4_ERR THEN
                GVL_SIG.G4_ERR := FALSE;
                GVL_SIG.G3_CODE_DEFAUT := 7; Step := 202; END_IF;
        14: GVL_SIG.G8_REQ        := TRUE;
            GVL_SIG.G8_ID_ATTENDU := GVL_MOULES.MOULE_DEMANDE;
            SubA := 15;
        15: IF GVL_SIG.G8_DONE THEN
                GVL_SIG.G8_DONE := FALSE;
                IF GVL_SIG.G8_OK THEN
                    GVL_MOULES.CH[GVL_MOULES.CIBLE_PRISE_CH,
                                  GVL_MOULES.CIBLE_PRISE_NV].RFID_OK := TRUE;
                    SubA := 16;
                ELSE
                    GVL_SIG.G8_ERR         := FALSE;
                    GVL_SIG.G3_CODE_DEFAUT := 8;
                    Step := 202;
                END_IF;
            ELSIF GVL_SIG.G8_ERR THEN
                GVL_SIG.G8_ERR         := FALSE;
                GVL_SIG.G3_CODE_DEFAUT := 8; Step := 202; END_IF;
        16: GVL_SIG.G5_REQ   := TRUE;
            GVL_SIG.G5_CIBLE := GVL_MOULES.CIBLE_PRISE_NV;
            SubA := 17;
        17: IF GVL_SIG.G5_DONE THEN
                GVL_SIG.G5_DONE := FALSE; SubA := 18;
            ELSIF GVL_SIG.G5_ERR THEN
                GVL_SIG.G5_ERR := FALSE;
                GVL_SIG.G3_CODE_DEFAUT := 6; Step := 202; END_IF;
        18: GVL_SIG.G7_REQ := TRUE;
            GVL_SIG.G7_CMD := 0; // EXT
            SubA := 19;
        19: IF GVL_SIG.G7_DONE THEN
                GVL_SIG.G7_DONE := FALSE; SubA := 20;
            ELSIF GVL_SIG.G7_ERR THEN
                GVL_SIG.G7_ERR := FALSE;
                GVL_SIG.G3_CODE_DEFAUT := 11; Step := 202; END_IF;
        20: GVL_SIG.G5_REQ   := TRUE;
            GVL_SIG.G5_CIBLE := 3; // Z_TRANSPORT
            SubA := 21;
        21: IF GVL_SIG.G5_DONE THEN
                GVL_SIG.G5_DONE := FALSE;
                IF NOT GVL_IO.CAPTEUR_CHARGE_CHARIOT THEN
                    GVL_SIG.G3_CODE_DEFAUT := 10; Step := 202;
                ELSE
                    SubA := 22;
                END_IF;
            ELSIF GVL_SIG.G5_ERR THEN
                GVL_SIG.G5_ERR := FALSE;
                GVL_SIG.G3_CODE_DEFAUT := 6; Step := 202; END_IF;
        22: GVL_SIG.G7_REQ := TRUE;
            GVL_SIG.G7_CMD := 1; // RET
            SubA := 23;
        23: IF GVL_SIG.G7_DONE THEN
                GVL_SIG.G7_DONE := FALSE;
                GVL_MOULES.CH[GVL_MOULES.CIBLE_PRISE_CH,
                               GVL_MOULES.CIBLE_PRISE_NV].OCCUPE := FALSE;
                GVL_MOULES.CH[GVL_MOULES.CIBLE_PRISE_CH,
                               GVL_MOULES.CIBLE_PRISE_NV].ID     := 0;
                GVL_MOULES.NB_EMPLACEMENTS_LIBRES :=
                    GVL_MOULES.NB_EMPLACEMENTS_LIBRES + 1;
                GVL_SEQ.MOULE_EN_TRANSIT := TRUE;
                SubA := 24;
            ELSIF GVL_SIG.G7_ERR THEN
                GVL_SIG.G7_ERR := FALSE;
                GVL_SIG.G3_CODE_DEFAUT := 11; Step := 203; END_IF;
        24: GVL_SIG.G4_REQ   := TRUE;
            GVL_SIG.G4_CIBLE := 0; // P0
            SubA := 25;
        25: IF GVL_SIG.G4_DONE THEN
                GVL_SIG.G4_DONE := FALSE; SubA := 26;
            ELSIF GVL_SIG.G4_ERR THEN
                GVL_SIG.G4_ERR := FALSE;
                GVL_SIG.G3_CODE_DEFAUT := 7; Step := 203; END_IF;
        26: GVL_SIG.G8_REQ        := TRUE;
            GVL_SIG.G8_ID_ATTENDU := GVL_MOULES.MOULE_DEMANDE;
            SubA := 27;
        27: IF GVL_SIG.G8_DONE THEN
                GVL_SIG.G8_DONE := FALSE;
                IF GVL_SIG.G8_OK THEN
                    BrA_Done := TRUE;
                ELSE
                    GVL_SIG.G8_ERR         := FALSE;
                    GVL_SIG.G3_CODE_DEFAUT := 9;
                    Step := 210;
                END_IF;
            ELSIF GVL_SIG.G8_ERR THEN
                GVL_SIG.G8_ERR         := FALSE;
                GVL_SIG.G3_CODE_DEFAUT := 9; Step := 210; END_IF;
        END_CASE;
    END_IF;

    IF NOT BrB_Done THEN
        CASE SubB OF
        0:  GVL_SIG.VYT_NETTOYAGE  := TRUE;
            GVL_IO.VOYANT_NETTOYAGE := TRUE;
            IF SubA >= 10 THEN
                GVL_IO.BUZZER_DEBUT_NETTOYAGE := TRUE;
                NettoyageTimerEnable := TRUE;
                ProlongTimerEnable := FALSE;
                GVL_SIG.NETTOYAGE_EN_COURS := TRUE;
                GVL_SIG.NETTOYAGE_TIMEOUT := FALSE;
                GVL_SIG.NETTOYAGE_PROLONGATION_UTILISEE := FALSE;
                GVL_SIG.NETTOYAGE_DEPASSEMENT_MAX := FALSE;
                SubB := 1;
            END_IF;

        1:  GVL_IO.BUZZER_DEBUT_NETTOYAGE := FALSE;
            GVL_SIG.VYT_ATTENTE_ZONE := NOT GVL_SIG.ZONE_CONFIRMEE;
            GVL_IO.VOYANT_ATTENTE_ZONE_LIBRE := NOT GVL_SIG.ZONE_CONFIRMEE;

            IF GVL_SIG.ZONE_CONFIRMEE THEN
                GVL_IO.VOYANT_NETTOYAGE := FALSE;
                GVL_IO.VOYANT_ATTENTE_ZONE_LIBRE := FALSE;
                GVL_IO.VOYANT_NETTOYAGE_TIMEOUT := FALSE;
                GVL_IO.VOYANT_NETTOYAGE_MAX := FALSE;
                GVL_IO.BUZZER_ATTENTE_ZONE_LIBRE := FALSE;
                GVL_SIG.VYT_NETTOYAGE := FALSE;
                GVL_SIG.VYT_ATTENTE_ZONE := FALSE;
                GVL_SIG.VYT_NETTOYAGE_TIMEOUT := FALSE;
                GVL_SIG.NETTOYAGE_EN_COURS := FALSE;
                GVL_SIG.NETTOYAGE_TIMEOUT := FALSE;
                NettoyageTimerEnable := FALSE;
                ProlongTimerEnable := FALSE;
                BrB_Done := TRUE;

            ELSIF T_Prolong5.Q THEN
                GVL_SIG.NETTOYAGE_DEPASSEMENT_MAX := TRUE;
                GVL_SIG.NETTOYAGE_TIMEOUT := TRUE;
                GVL_SIG.VYT_NETTOYAGE_TIMEOUT := TRUE;
                GVL_IO.VOYANT_NETTOYAGE_TIMEOUT := TRUE;
                GVL_IO.VOYANT_NETTOYAGE_MAX := TRUE;
                GVL_IO.BUZZER_ATTENTE_ZONE_LIBRE := TRUE;
                GVL_SIG.G3_CODE_DEFAUT := 18;
                IF GVL_SEQ.MOULE_EN_TRANSIT THEN
                    Step := 203;
                ELSE
                    Step := 202;
                END_IF;

            ELSIF T_Nettoyage15.Q THEN
                GVL_SIG.NETTOYAGE_TIMEOUT := TRUE;
                GVL_SIG.VYT_NETTOYAGE_TIMEOUT := TRUE;
                GVL_IO.VOYANT_NETTOYAGE_TIMEOUT := TRUE;
                GVL_IO.BUZZER_ATTENTE_ZONE_LIBRE := TRUE;

                IF GVL_SIG.OP_PROLONG_NETTOYAGE
                   AND NOT GVL_SIG.NETTOYAGE_PROLONGATION_UTILISEE THEN
                    GVL_SIG.NETTOYAGE_PROLONGATION_UTILISEE := TRUE;
                    GVL_SIG.NETTOYAGE_TIMEOUT := FALSE;
                    GVL_SIG.VYT_NETTOYAGE_TIMEOUT := FALSE;
                    GVL_IO.VOYANT_NETTOYAGE_TIMEOUT := FALSE;
                    GVL_IO.BUZZER_ATTENTE_ZONE_LIBRE := FALSE;
                    NettoyageTimerEnable := FALSE;
                    ProlongTimerEnable := TRUE;
                END_IF;
            END_IF;
        END_CASE;
    END_IF;

    IF BrA_Done AND BrB_Done THEN
        Step := 30;
    END_IF;

// ════════════════════════════════════════════════════════════
// PHASE 3 — Dépôt nouveau moule sur introducteur
// ════════════════════════════════════════════════════════════
30:
    GVL_SIG.G6_REQ   := TRUE;
    GVL_SIG.G6_CIBLE := 0; // NORD
    Step := 31;

31:
    IF GVL_SIG.G6_DONE THEN
        GVL_SIG.G6_DONE := FALSE; Step := 32;
    ELSIF GVL_SIG.G6_ERR THEN
        GVL_SIG.G6_ERR         := FALSE;
        GVL_SIG.G3_CODE_DEFAUT := 11; Step := 203; END_IF;

32:
    GVL_SIG.G7_REQ := TRUE;
    GVL_SIG.G7_CMD := 0; // EXT
    Step := 33;

33:
    IF GVL_SIG.G7_DONE THEN
        GVL_SIG.G7_DONE := FALSE; Step := 34;
    ELSIF GVL_SIG.G7_ERR THEN
        GVL_SIG.G7_ERR         := FALSE;
        GVL_SIG.G3_CODE_DEFAUT := 11; Step := 203; END_IF;

34:
    GVL_SIG.G5_REQ   := TRUE;
    GVL_SIG.G5_CIBLE := 0; // Z_ZPM
    Step := 35;

35:
    IF GVL_SIG.G5_DONE THEN
        GVL_SIG.G5_DONE := FALSE; Step := 36;
    ELSIF GVL_SIG.G5_ERR THEN
        GVL_SIG.G5_ERR         := FALSE;
        GVL_SIG.G3_CODE_DEFAUT := 6; Step := 203; END_IF;

36:
    GVL_SIG.G7_REQ := TRUE;
    GVL_SIG.G7_CMD := 1; // RET
    Step := 37;

37:
    IF GVL_SIG.G7_DONE THEN
        GVL_SIG.G7_DONE := FALSE;
        IF NOT GVL_IO.MOULE_SUR_INTRO THEN
            GVL_SIG.G3_CODE_DEFAUT := 11; Step := 203;
        ELSIF GVL_IO.CAPTEUR_CHARGE_CHARIOT THEN
            GVL_SIG.G3_CODE_DEFAUT := 11; Step := 203;
        ELSE
            Step := 38;
        END_IF;
    ELSIF GVL_SIG.G7_ERR THEN
        GVL_SIG.G7_ERR         := FALSE;
        GVL_SIG.G3_CODE_DEFAUT := 11; Step := 203; END_IF;

38:
    GVL_SIG.G5_REQ   := TRUE;
    GVL_SIG.G5_CIBLE := 3; // Z_TRANSPORT
    Step := 39;

39:
    IF GVL_SIG.G5_DONE THEN
        GVL_SIG.G5_DONE         := FALSE;
        GVL_SIG.G10_REQ_ENTRER  := TRUE;
        GVL_SIG.G9_REQ_BRIDAGE  := TRUE;
        Step := 40;
    ELSIF GVL_SIG.G5_ERR THEN
        GVL_SIG.G5_ERR         := FALSE;
        GVL_SIG.G3_CODE_DEFAUT := 6; Step := 203; END_IF;

40:
    IF GVL_SIG.G9_BRIDE_OK AND GVL_SIG.G10_A_ZPM THEN
        GVL_MOULES.MOULE_EN_PRESSE := GVL_MOULES.MOULE_DEMANDE;
        GVL_SEQ.MOULE_EN_TRANSIT   := FALSE;
        GVL_SIG.G10_REQ_ENTRER     := FALSE;
        Step := 41;
    ELSIF GVL_SIG.G9_DEFAUT THEN
        GVL_SIG.G3_CODE_DEFAUT := 3; Step := 200;
    ELSIF GVL_SIG.G10_DEFAUT THEN
        GVL_SIG.G3_CODE_DEFAUT := 5; Step := 200;
    END_IF;

// ════════════════════════════════════════════════════════════
// DIVERGENCE ET#3 — Autorisation presse ‖ Retour garage
// ════════════════════════════════════════════════════════════
41:
    BrA_Done := FALSE;
    BrB_Done := FALSE;
    SubA     := 0;
    SubB     := 0;
    Step     := 42;

42:
    IF NOT BrA_Done THEN
        CASE SubA OF
        0:  GVL_SIG.G9_REQ_AUTORISER := TRUE;
            SubA := 1;
        1:  IF GVL_SIG.G9_AUTORISE_OK THEN
                GVL_SIG.G9_REQ_AUTORISER := FALSE;
                BrA_Done := TRUE;
            ELSIF GVL_SIG.G9_DEFAUT THEN
                GVL_SIG.G3_CODE_DEFAUT := 3; Step := 200; END_IF;
        END_CASE;
    END_IF;

    IF NOT BrB_Done THEN
        CASE SubB OF
        0:  GVL_SIG.G4_REQ   := TRUE;
            GVL_SIG.G4_CIBLE := 6; // P6 Garage
            SubB := 1;
        1:  IF GVL_SIG.G4_DONE THEN
                GVL_SIG.G4_DONE := FALSE;
                BrB_Done := TRUE;
            ELSIF GVL_SIG.G4_ERR THEN
                GVL_SIG.G4_ERR := FALSE;
                BrB_Done := TRUE;  // Non bloquant
            END_IF;
        END_CASE;
    END_IF;

    IF BrA_Done AND BrB_Done THEN
        Step := 50;
    END_IF;

// ════════════════════════════════════════════════════════════
// PHASE FINALE — Fin de cycle
// ════════════════════════════════════════════════════════════
50:
    GVL_SEQ.CYCLE_INTERROMPU    := FALSE;
    GVL_SEQ.CYCLE_EN_COURS      := FALSE;
    GVL_MOULES.ALM_STOCK_PLEIN  := FALSE;
    GVL_SIG.VYT_CYCLE_EN_COURS  := FALSE;
    GVL_SIG.G3_FIN_CM           := TRUE;
    IF NOT GVL_SIG.G3_REQ THEN
        GVL_SIG.G3_FIN_CM := FALSE;
        Step := 0;
    END_IF;

// ════════════════════════════════════════════════════════════
// BRANCHES DÉFAUT
// ════════════════════════════════════════════════════════════
200: // Défaut chariot VIDE
    GVL_SIG.G3_DEFAUT          := TRUE;
    GVL_SEQ.DEFAUT_ACTIF       := TRUE;
    GVL_SEQ.CODE_DEFAUT        := GVL_SIG.G3_CODE_DEFAUT;
    GVL_SIG.VYT_CYCLE_EN_COURS := FALSE;
    GVL_SIG.VYT_DEFAUT         := TRUE;
    IF GVL_MOULES.CIBLE_DEPOT_CH >= 1
       AND GVL_MOULES.CIBLE_DEPOT_CH <= 5 THEN
        GVL_MOULES.CH[GVL_MOULES.CIBLE_DEPOT_CH,
                      GVL_MOULES.CIBLE_DEPOT_NV].RESERVE := FALSE;
    END_IF;
    IF GVL_SIG.OP_CMD_RESET AND GVL_SIG.OP_CMD_ACQ THEN
        GVL_SIG.G3_DEFAUT    := FALSE;
        GVL_SEQ.DEFAUT_ACTIF := FALSE;
        GVL_SEQ.CODE_DEFAUT  := 0;
        GVL_SIG.VYT_DEFAUT   := FALSE;
        GVL_SEQ.CYCLE_INTERROMPU := FALSE;
        Step := 0;
    END_IF;

201: // Défaut ancien moule sur fourches
    GVL_SIG.G3_DEFAUT          := TRUE;
    GVL_SEQ.DEFAUT_ACTIF       := TRUE;
    GVL_SEQ.CODE_DEFAUT        := GVL_SIG.G3_CODE_DEFAUT;
    GVL_SIG.VYT_DEFAUT         := TRUE;
    GVL_SIG.VYT_CYCLE_EN_COURS := FALSE;
    IF GVL_SIG.OP_CMD_RESET AND GVL_SIG.OP_CMD_ACQ THEN
        GVL_SIG.G3_DEFAUT    := FALSE;
        GVL_SEQ.DEFAUT_ACTIF := FALSE;
        GVL_SIG.VYT_DEFAUT   := FALSE;
        Step := 0;
    END_IF;

202: // Défaut ancien moule déposé, chariot vide
    GVL_SIG.G3_DEFAUT          := TRUE;
    GVL_SEQ.DEFAUT_ACTIF       := TRUE;
    GVL_SEQ.CODE_DEFAUT        := GVL_SIG.G3_CODE_DEFAUT;
    GVL_SIG.VYT_DEFAUT         := TRUE;
    GVL_SIG.VYT_CYCLE_EN_COURS := FALSE;
    IF GVL_SIG.OP_CMD_RESET AND GVL_SIG.OP_CMD_ACQ THEN
        GVL_SIG.G3_DEFAUT    := FALSE;
        GVL_SEQ.DEFAUT_ACTIF := FALSE;
        GVL_SIG.VYT_DEFAUT   := FALSE;
        Step := 0;
    END_IF;

203: // Défaut nouveau moule sur fourches (MOULE_EN_TRANSIT=TRUE)
    GVL_SIG.G3_DEFAUT          := TRUE;
    GVL_SEQ.DEFAUT_ACTIF       := TRUE;
    GVL_SEQ.CODE_DEFAUT        := GVL_SIG.G3_CODE_DEFAUT;
    GVL_SIG.VYT_DEFAUT         := TRUE;
    GVL_SIG.VYT_CYCLE_EN_COURS := FALSE;
    IF GVL_SIG.OP_CMD_RESET AND GVL_SIG.OP_CMD_ACQ THEN
        GVL_SIG.G3_DEFAUT    := FALSE;
        GVL_SEQ.DEFAUT_ACTIF := FALSE;
        GVL_SIG.VYT_DEFAUT   := FALSE;
        Step := 0;
    END_IF;

210: // RFID2 KO — ROLLBACK (remettre moule en chambre prise)
    GVL_SIG.ALM_RFID           := TRUE;
    GVL_SIG.G3_DEFAUT          := TRUE;
    GVL_SEQ.DEFAUT_ACTIF       := TRUE;
    GVL_SEQ.CODE_DEFAUT        := 9;
    GVL_SIG.VYT_CYCLE_EN_COURS := FALSE;
    GVL_SIG.VYT_DEFAUT         := TRUE;
    GVL_MOULES.CH[GVL_MOULES.CIBLE_PRISE_CH,
                  GVL_MOULES.CIBLE_PRISE_NV].OCCUPE := TRUE;
    GVL_MOULES.CH[GVL_MOULES.CIBLE_PRISE_CH,
                  GVL_MOULES.CIBLE_PRISE_NV].ID     := GVL_MOULES.MOULE_DEMANDE;
    GVL_MOULES.NB_EMPLACEMENTS_LIBRES :=
        GVL_MOULES.NB_EMPLACEMENTS_LIBRES - 1;
    GVL_SEQ.MOULE_EN_TRANSIT := FALSE;
    IF GVL_SIG.OP_CMD_RESET AND GVL_SIG.OP_CMD_ACQ THEN
        GVL_SIG.G3_DEFAUT    := FALSE;
        GVL_SEQ.DEFAUT_ACTIF := FALSE;
        GVL_SIG.ALM_RFID     := FALSE;
        GVL_SIG.VYT_DEFAUT   := FALSE;
        Step := 0;
    END_IF;

END_CASE;

END_FUNCTION_BLOCK

(* ---- 23_FB_HMI_Controller.st ---- *)
// ================================================================
// 23_FB_HMI_Controller.st  —  Contrôleur IHM CODESYS Visualization
// CODESYS V3.5 — FUNCTION_BLOCK
//
// Rôle :
//   - Génère les textes et couleurs dynamiques affichés dans la Visualization
//   - Détecte les fronts montants des boutons HMI (R_TRIG)
//   - Route les commandes HMI vers GVL_IO (puis → GVL_SIG via PRG_MAIN)
//   - Gère le chronomètre cycle et la barre de progression G3
//
// Appel dans PRG_MAIN : avant le bloc de copies GVL_IO → GVL_SIG
//
// Modification v2 — Laser OSSD :
//   - HMI_BTN_ZONE_OK supprimé du flux normal (ZONE_CONFIRMEE géré par FB_LaserSafe)
//   - rZoneOk supprimé
// ================================================================

FUNCTION_BLOCK FB_HMI_Controller
VAR
    // ── Fronts montants boutons ───────────────────────────────────
    rHoming   : R_TRIG;
    rCmdCM    : R_TRIG;
    rAcq      : R_TRIG;

    // ── Chronomètre cycle ─────────────────────────────────────────
    tTick       : TON;
    iCycleSec   : DINT;
    bCycleWas   : BOOL;
    iMin, iSec  : DINT;
    sMin, sSec  : STRING(3);

    // ── Boucle stock ──────────────────────────────────────────────
    iCh, iNv    : INT;
END_VAR

// ── 1. MODE SYSTÈME → texte + couleur ────────────────────────────
IF GVL_SIG.OP_AU THEN
    GVL_HMI.HMI_MODE_TXT := 'ARRET URGENCE';
    GVL_HMI.HMI_COL_MODE := 16#FFFF3030;   // rouge vif
ELSIF GVL_SEQ.DEFAUT_ACTIF THEN
    GVL_HMI.HMI_MODE_TXT := 'DEFAUT';
    GVL_HMI.HMI_COL_MODE := 16#FFFF6600;   // orange défaut
ELSIF GVL_SEQ.CYCLE_EN_COURS THEN
    GVL_HMI.HMI_MODE_TXT := 'CYCLE EN COURS';
    GVL_HMI.HMI_COL_MODE := 16#FF00C800;   // vert cycle
ELSIF GVL_SEQ.HOMING_OK AND GVL_SIG.VYT_MACHINE_PRETE THEN
    GVL_HMI.HMI_MODE_TXT := 'EN ATTENTE';
    GVL_HMI.HMI_COL_MODE := 16#FF1C6EBF;   // bleu attente
ELSIF GVL_SIG.G2_REQ THEN
    GVL_HMI.HMI_MODE_TXT := 'HOMING...';
    GVL_HMI.HMI_COL_MODE := 16#FFFFA500;   // orange homing
ELSE
    GVL_HMI.HMI_MODE_TXT := 'HORS SERVICE';
    GVL_HMI.HMI_COL_MODE := 16#FF404040;   // gris
END_IF;

// ── 2. MOULE EN PRESSE → texte ────────────────────────────────────
GVL_HMI.HMI_MOULE_PRESSE_TXT := FC_MouleIDToStr(GVL_MOULES.MOULE_EN_PRESSE);

// ── 3. STOCK 5×2 → tableau de textes ─────────────────────────────
FOR iCh := 1 TO 5 DO
    FOR iNv := 1 TO 2 DO
        GVL_HMI.HMI_STOCK_TXT[iCh, iNv] := FC_MouleIDToStr(GVL_MOULES.CH[iCh, iNv].ID);
    END_FOR;
END_FOR;

// ── 4. PROGRESSION G3 ─────────────────────────────────────────────
GVL_HMI.HMI_G3_ETAPE    := GVL_SEQ.ETAPE_ACTIVE;
GVL_HMI.HMI_ETAPE_G3_TXT := FC_EtapeG3ToStr(GVL_SEQ.ETAPE_ACTIVE);
IF GVL_SEQ.CYCLE_EN_COURS AND GVL_SEQ.ETAPE_ACTIVE > 0 THEN
    GVL_HMI.HMI_G3_PCT := INT_TO_REAL(GVL_SEQ.ETAPE_ACTIVE) * 100.0 / 15.0;
ELSE
    GVL_HMI.HMI_G3_PCT := 0.0;
END_IF;

// ── 5. CHRONOMÈTRE CYCLE ──────────────────────────────────────────
IF GVL_SEQ.CYCLE_EN_COURS AND NOT bCycleWas THEN
    iCycleSec := 0;
    bCycleWas := TRUE;
ELSIF NOT GVL_SEQ.CYCLE_EN_COURS THEN
    bCycleWas := FALSE;
    tTick(IN := FALSE);
END_IF;
IF GVL_SEQ.CYCLE_EN_COURS THEN
    tTick(IN := TRUE, PT := T#1S);
    IF tTick.Q THEN
        iCycleSec := iCycleSec + 1;
        tTick(IN := FALSE);
    END_IF;
END_IF;
iMin := iCycleSec / 60;
iSec := iCycleSec MOD 60;
IF iMin < 10 THEN sMin := CONCAT('0', DINT_TO_STRING(iMin));
ELSE sMin := DINT_TO_STRING(iMin); END_IF;
IF iSec < 10 THEN sSec := CONCAT('0', DINT_TO_STRING(iSec));
ELSE sSec := DINT_TO_STRING(iSec); END_IF;
GVL_HMI.HMI_TEMPS_CYCLE := CONCAT(sMin, CONCAT(':', sSec));

// ── 6. SÉLECTEUR MOULE ────────────────────────────────────────────
GVL_HMI.HMI_SEL_MOULE_OK := (GVL_HMI.HMI_SEL_MOULE >= 1)
                          AND (GVL_HMI.HMI_SEL_MOULE <= 5);

// ── 7. BOUTONS → GVL_IO (détection front montant) ─────────────────

// HOMING
rHoming(CLK := GVL_HMI.HMI_BTN_HOMING);
IF rHoming.Q THEN
    GVL_IO.CMD_HOMING_MANUEL := TRUE;
ELSIF NOT GVL_SIG.G2_REQ THEN
    GVL_IO.CMD_HOMING_MANUEL := FALSE;
END_IF;

// ACQUITTEMENT DÉFAUTS
rAcq(CLK := GVL_HMI.HMI_BTN_ACQ);
IF rAcq.Q THEN
    GVL_IO.CMD_ACQ_DEF := TRUE;
ELSE
    GVL_IO.CMD_ACQ_DEF := FALSE;
END_IF;

// ZONE LIBRE : désormais pilotée automatiquement par FB_LaserSafe (OSSD Sick S3000)
// HMI_BTN_ZONE_OK conservé dans GVL_HMI uniquement pour diagnostic Visualization
// (ne déclenche plus ZONE_CONFIRMEE en production — laser prime)

// ARRÊT URGENCE SW
GVL_IO.AU_ACTIF := GVL_HMI.HMI_BTN_AU;

// CMD_CM — ne démarre que si un moule valide est sélectionné
rCmdCM(CLK := GVL_HMI.HMI_BTN_CMD_CM);
IF rCmdCM.Q AND GVL_HMI.HMI_SEL_MOULE_OK THEN
    GVL_IO.MOULE_DEMANDE_HMI := INT_TO_USINT(GVL_HMI.HMI_SEL_MOULE);
    GVL_IO.CMD_CM := TRUE;
ELSIF NOT GVL_SEQ.CYCLE_EN_COURS THEN
    GVL_IO.CMD_CM := FALSE;
END_IF;

// ── 8. INDICATEUR ALARME GLOBALE ─────────────────────────────────
GVL_HMI.HMI_ALARME_ACTIVE :=
    GVL_SIG.ALM_STOCK_PLEIN   OR GVL_SIG.ALM_RFID        OR
    GVL_SIG.ALM_DEBRIDAGE      OR GVL_SIG.ALM_BRIDAGE      OR
    GVL_SIG.ALM_PILON          OR GVL_SIG.ALM_INTRO        OR
    GVL_SIG.ALM_AXE_X          OR GVL_SIG.ALM_AXE_Z        OR
    GVL_SIG.ALM_ROTATION       OR GVL_SIG.ALM_SATELLITE     OR
    GVL_SIG.ALM_COMM_PRESSE    OR GVL_SIG.ALM_ZONE         OR
    GVL_SIG.ALM_HOMING;

(* ---- 24_FB_FaultInjector.st ---- *)
// ================================================================
// 24_FB_FaultInjector.st  —  Injection scénarios modes dégradés
// CODESYS V3.5 — FUNCTION_BLOCK
//
// Utilisé UNIQUEMENT en mode simulation/soutenance pour démontrer
// la réaction du système aux 8 modes dégradés du cahier des charges.
//
// Appelé par FB_HMI_Controller via la Visualization (écran 4)
//
// IMPORTANT : ResetFlt remet toutes les variables à leur état normal
// ================================================================

FUNCTION_BLOCK FB_FaultInjector
VAR_INPUT
    FaultID   : INT;    // 0-8 : scénario sélectionné
    Inject    : BOOL;   // R_TRIG depuis bouton INJECTER
    ResetFlt  : BOOL;   // R_TRIG depuis bouton RESET
END_VAR
VAR_OUTPUT
    Desc      : STRING(100);  // Description affichée avant injection
    Result    : STRING(120);  // Résultat affiché après injection
    FltActive : BOOL;         // TRUE si défaut injecté en cours
END_VAR
VAR
    bInjected   : BOOL;           // défaut actuellement injecté
    iInjectedID : INT;            // ID du défaut injecté
    tAutoReset  : TON;            // timeout auto-reset pour D3, D4
    rInj        : R_TRIG;
    rRst        : R_TRIG;
END_VAR

// ── Détection fronts ──────────────────────────────────────────────
rInj(CLK := Inject);
rRst(CLK := ResetFlt);

// ── Description (mise à jour à chaque cycle selon sélection) ──────
IF NOT bInjected THEN
    CASE FaultID OF
        0: Desc := 'Sélectionner un scénario de défaut...';
        1: Desc := 'D1 — Stock plein : aucune chambre libre. G3 refuse le démarrage.';
        2: Desc := 'D2 — Moule absent : ID demandé introuvable en stock.';
        3: Desc := 'D3 — Timeout axe X : déplacement bloqué (simulé).';
        4: Desc := 'D4 — RFID KO : 3 tentatives échouées, rollback moule.';
        5: Desc := 'D5 — Cycle interrompu : simule coupure secteur en cours de cycle.';
        6: Desc := 'D6 — Zone opérateurs : zone non libérée, cycle bloqué en S14.';
        7: Desc := 'D7 — Perte Profinet : presse inaccessible, arrêt tous mouvements.';
        8: Desc := 'D8 — Coupure secteur : AU + CYCLE_INTERROMPU retain, homing obligatoire.';
    ELSE
        Desc := '???';
    END_CASE;
END_IF;

// ── INJECTION ─────────────────────────────────────────────────────
IF rInj.Q AND NOT bInjected AND FaultID >= 1 AND FaultID <= 8 THEN
    bInjected   := TRUE;
    iInjectedID := FaultID;
    tAutoReset(IN := FALSE);

    CASE FaultID OF

        1: // D1 — Stock plein
            GVL_MOULES.NB_EMPLACEMENTS_LIBRES := 0;
            // Forcer toutes les chambres occupées
            GVL_MOULES.CH[5,1].OCCUPE := TRUE;
            GVL_MOULES.CH[5,2].OCCUPE := TRUE;
            Result := 'D1 injecté : NB_EMPLACEMENTS_LIBRES=0. Appuyez CMD_CM → alarme ALM_STOCK_PLEIN attendue.';

        2: // D2 — Moule absent
            GVL_IO.MOULE_DEMANDE_HMI := 9;   // ID 9 n'existe pas en stock
            GVL_MOULES.MOULE_DEMANDE := 9;
            Result := 'D2 injecté : MOULE_DEMANDE=ID9 (inexistant). Appuyez CMD_CM → G3 ne démarre pas.';

        3: // D3 — Timeout axe X (injecter erreur axe X)
            GVL_SIG.G4_ERR := TRUE;
            Result := 'D3 injecté : G4_ERR=TRUE. Si cycle en cours → G3 défaut, alarme ALM_AXE_X.';
            tAutoReset(IN := TRUE, PT := T#10S);  // auto-clear après 10s

        4: // D4 — RFID KO
            GVL_SIG.G8_ERR := TRUE;
            GVL_SIG.G8_OK  := FALSE;
            Result := 'D4 injecté : G8_ERR=TRUE. Si cycle en cours → 3 tentatives RFID → rollback → G3 défaut.';
            tAutoReset(IN := TRUE, PT := T#10S);

        5: // D5 — Cycle interrompu (simule coupure secteur)
            GVL_SEQ.CYCLE_INTERROMPU := TRUE;
            GVL_IO.AU_ACTIF := TRUE;
            Result := 'D5 injecté : CYCLE_INTERROMPU=TRUE + AU. Au reset : G0 passe en E2 (alarme reprise), homing obligatoire.';

        6: // D6 — Zone opérateurs
            GVL_IO.CAPTEUR_ZONE_OCCUPEE := TRUE;
            GVL_SIG.ZONE_CONFIRMEE := FALSE;
            GVL_HMI.HMI_BTN_ZONE_OK := FALSE;
            Result := 'D6 injecté : Zone occupée + ZONE_CONFIRMEE=FALSE. Cycle bloqué en S14 → voyant nettoyage actif.';

        7: // D7 — Perte Profinet
            GVL_SIG.PERTE_PROFINET := TRUE;
            GVL_SIG.ALM_COMM_PRESSE := TRUE;
            Result := 'D7 injecté : PERTE_PROFINET=TRUE. G9 ne peut pas commander la presse → arrêt général.';

        8: // D8 — Coupure secteur
            GVL_IO.AU_ACTIF := TRUE;
            GVL_SEQ.CYCLE_INTERROMPU := TRUE;
            GVL_SEQ.MOULE_EN_TRANSIT := TRUE;
            Result := 'D8 injecté : AU + CYCLE_INTERROMPU + MOULE_EN_TRANSIT. Redémarrer → G0 exige homing + acquittement.';

    END_CASE;
END_IF;

// ── Auto-reset D3/D4 après timeout ───────────────────────────────
tAutoReset(IN := bInjected AND (iInjectedID = 3 OR iInjectedID = 4));
IF tAutoReset.Q THEN
    GVL_SIG.G4_ERR := FALSE;
    GVL_SIG.G8_ERR := FALSE;
    GVL_SIG.G8_OK  := FALSE;
    bInjected   := FALSE;
    iInjectedID := 0;
    Result := 'Auto-reset D3/D4 effectué après 10s.';
    tAutoReset(IN := FALSE);
END_IF;

// ── RESET MANUEL ──────────────────────────────────────────────────
IF rRst.Q THEN
    // Remettre toutes les variables injectées à leur état normal
    GVL_MOULES.NB_EMPLACEMENTS_LIBRES := 4;  // 4 emplacements libres par défaut
    GVL_MOULES.CH[5,1].OCCUPE := FALSE;
    GVL_MOULES.CH[5,2].OCCUPE := FALSE;
    GVL_IO.MOULE_DEMANDE_HMI := 0;
    GVL_MOULES.MOULE_DEMANDE := 0;
    GVL_SIG.G4_ERR := FALSE;
    GVL_SIG.G8_ERR := FALSE;
    GVL_SIG.G8_OK  := FALSE;
    GVL_SEQ.CYCLE_INTERROMPU := FALSE;
    GVL_SEQ.MOULE_EN_TRANSIT := FALSE;
    GVL_IO.AU_ACTIF := FALSE;
    GVL_HMI.HMI_BTN_AU := FALSE;
    GVL_IO.CAPTEUR_ZONE_OCCUPEE := FALSE;
    GVL_SIG.PERTE_PROFINET := FALSE;
    GVL_SIG.ALM_COMM_PRESSE := FALSE;
    // Acquitter alarmes
    GVL_SIG.ALM_STOCK_PLEIN  := FALSE;
    GVL_SIG.ALM_RFID         := FALSE;
    GVL_SIG.ALM_AXE_X        := FALSE;
    GVL_SIG.ALM_AXE_Z        := FALSE;
    GVL_SIG.ALM_ZONE         := FALSE;
    GVL_SIG.ALM_HOMING       := FALSE;
    GVL_SEQ.DEFAUT_ACTIF     := FALSE;
    GVL_SEQ.CODE_DEFAUT      := 0;
    bInjected   := FALSE;
    iInjectedID := 0;
    tAutoReset(IN := FALSE);
    Result   := 'Reset complet effectué. Système remis à l état nominal.';
    Desc     := 'Sélectionner un scénario de défaut...';
END_IF;

FltActive := bInjected;
GVL_HMI.HMI_FAULT_ACTIVE := bInjected;

// Couleur bouton INJECTER : rouge foncé si déjà actif, rouge vif sinon
IF bInjected THEN
    GVL_HMI.HMI_COL_FAULT_BTN := 16#FF8B0000;   // rouge foncé = déjà injecté
ELSE
    GVL_HMI.HMI_COL_FAULT_BTN := 16#FFCC0000;   // rouge vif = prêt à injecter
END_IF;

(* ---- 25_FB_LaserSafe.st ---- *)
// ================================================================
// 25_FB_LaserSafe.st  —  Gestion barrière laser 2D (Sick S3000 OSSD)
// CODESYS V3.5 — FUNCTION_BLOCK
//
// Rôle :
//   Remplace le bouton ZONE_LIBRE (ZONE_LIBRE_BTN) par une validation
//   automatique basée sur les sorties OSSD des scanners 2D.
//
//   Logique :
//     1. Lecture OSSD_ZPM et OSSD_PRESSE (TRUE = zone libre)
//     2. Muting automatique si CAPTEUR_Z_TRANSPORT = TRUE
//        (chariot en position haute — le faisceau serait déclenché
//         par le chariot lui-même lors du retour avec nouveau moule)
//     3. Timer T_Confirm = T_ZONE_LIBRE_CONFIRM (défaut T#10S)
//        Les deux zones doivent être libres en continu pendant 10s
//     4. Après 10s confirmées → OSSD_ZONE_LIBRE_AUTO := TRUE
//                              → ZONE_CONFIRMEE := TRUE
//     5. Ré-intrusion après validation → invalidation + alarme
//
// Appel dans PRG_MAIN : avant instG3 (coordinateur cycle)
// ================================================================

FUNCTION_BLOCK FB_LaserSafe
VAR
    T_Confirm      : TON;       // Timer confirmation 10s zone libre
    ConfirmTimerEN : BOOL;      // Enable timer
END_VAR

// ─── Muting automatique ───────────────────────────────────────────────────────
// Lorsque le chariot est en Z_TRANSPORT (hauteur de transit, bras levés),
// les lasers sont mutés pour éviter un faux déclenchement lors du retour
// chariot avec le nouveau moule.
GVL_SIG.LASER_MUTING_ACTIF := GVL_IO.CAPTEUR_Z_TRANSPORT;

// ─── Lecture OSSD (copie dans signaux inter-GRAFCETs) ────────────────────────
GVL_SIG.LASER_ZPM_LIBRE    := GVL_IO.OSSD_ZPM;
GVL_SIG.LASER_PRESSE_LIBRE := GVL_IO.OSSD_PRESSE;

// ─── Timer de confirmation 10s ────────────────────────────────────────────────
// Active uniquement si :
//   • les deux zones OSSD sont libres (= vraies)
//   • le muting n'est pas actif (chariot pas en transit)
//   • le nettoyage est en cours (phase ET#2 active)
//   • ZONE_CONFIRMEE pas encore validée (évite re-triggering)
ConfirmTimerEN :=  GVL_SIG.LASER_ZPM_LIBRE
               AND GVL_SIG.LASER_PRESSE_LIBRE
               AND NOT GVL_SIG.LASER_MUTING_ACTIF
               AND GVL_SIG.NETTOYAGE_EN_COURS
               AND NOT GVL_SIG.ZONE_CONFIRMEE;

T_Confirm(IN := ConfirmTimerEN, PT := GVL_CFG.T_ZONE_LIBRE_CONFIRM);

GVL_SIG.LASER_CONFIRM_EN_COURS := ConfirmTimerEN AND NOT T_Confirm.Q;

// ─── Confirmation automatique ─────────────────────────────────────────────────
// Quand le timer expire : zones libres depuis 10s → autoriser retour chariot
IF T_Confirm.Q THEN
    GVL_SIG.OSSD_ZONE_LIBRE_AUTO := TRUE;
    GVL_SIG.ZONE_CONFIRMEE       := TRUE;
END_IF;

// ─── Reset OSSD_ZONE_LIBRE_AUTO si conditions perdues ────────────────────────
// (avant validation — après, seul G3 reset ZONE_CONFIRMEE via ré-intrusion)
IF NOT ConfirmTimerEN AND GVL_SIG.NETTOYAGE_EN_COURS AND NOT GVL_SIG.ZONE_CONFIRMEE THEN
    GVL_SIG.OSSD_ZONE_LIBRE_AUTO := FALSE;
END_IF;

// ─── Ré-intrusion APRÈS validation ───────────────────────────────────────────
// Quelqu'un entre dans la zone après validation laser mais avant que le
// chariot soit revenu (LASER_MUTING_ACTIF indique le retour chariot en cours).
// → Invalider la validation et attendre une nouvelle confirmation 10s.
// → Déclencher alarme ALM_ZONE.
IF GVL_SIG.ZONE_CONFIRMEE
   AND GVL_SIG.NETTOYAGE_EN_COURS
   AND NOT GVL_SIG.LASER_MUTING_ACTIF
   AND (NOT GVL_IO.OSSD_ZPM OR NOT GVL_IO.OSSD_PRESSE) THEN
    GVL_SIG.ZONE_CONFIRMEE       := FALSE;
    GVL_SIG.OSSD_ZONE_LIBRE_AUTO := FALSE;
    GVL_SIG.ALM_ZONE             := TRUE;
END_IF;

END_FUNCTION_BLOCK
